(* IEC 61131-3 sources: daoli-st-library/DL_Process (part 15) *)

(* ---- FC_DL_PaddingPickupCalc.st ---- *)
(*
  DL Factory R83 | FC_DL_PaddingPickupCalc
  功能：由轧车前干重与轧后湿重算轧余率，并按克重门幅速度换算带液量。
  开源溯源：无（clean-room 自研，依据公开工艺公式，来源=行业通用公式，许可证=MIT，借鉴点=公式结构）
  规则：R1-R21 全遵守
*)
FUNCTION FC_DL_PaddingPickupCalc : REAL
VAR_INPUT
    fWetMassG : REAL; // 轧后湿重试样质量 [g] / Wet mass after padding [g]
    fDryMassG : REAL; // 轧前干重试样质量 [g] / Dry mass before padding [g]
    fSpeedMpm : REAL; // 轧车线速度 [m/min] / Padder line speed [m/min]
    fWidthM   : REAL; // 织物门幅 [m] / Fabric width [m]
    fGsm      : REAL; // 织物干克重 [g/m²] / Dry grammage [g/m^2]
END_VAR
VAR_OUTPUT
    fPickupPct : REAL; // 轧余率（带液量占干布重）[%] / Wet pickup [%]
    fCarryLpm  : REAL; // 每分钟带液量（密度按 1 kg/L 近似）[L/min] / Liquor carry-over [L/min]
    fCarryKgH  : REAL; // 每小时带液量 [kg/h] / Liquor carry-over [kg/h]
    xValid     : BOOL; // 计算有效性标志 / Calculation validity flag
END_VAR
VAR
    fDryKgMin : REAL; // 每分钟干布质量 [kg/min] / Dry fabric mass per minute [kg/min]
END_VAR
// 出口预置：四出口统一预置（R256）
fPickupPct := 0.0; fCarryLpm := 0.0; fCarryKgH := 0.0; xValid := FALSE;
// 非有限拦截 + 量纲自检 + 湿干重次序闸（R20/R21）
IF NOT (fWetMassG > -1.0E30 AND fWetMassG < 1.0E30) OR NOT (fDryMassG > -1.0E30 AND fDryMassG < 1.0E30) OR NOT (fSpeedMpm > -1.0E30 AND fSpeedMpm < 1.0E30) OR NOT (fWidthM > -1.0E30 AND fWidthM < 1.0E30) OR NOT (fGsm > -1.0E30 AND fGsm < 1.0E30) OR fDryMassG <= 0.0 OR fSpeedMpm <= 0.0 OR fWidthM <= 0.0 OR fGsm <= 0.0 OR fWetMassG < fDryMassG THEN
    FC_DL_PaddingPickupCalc := -1.0; RETURN;   // 哨兵 -1：非有限或量纲/次序越界 / Sentinel -1
END_IF
// 轧余率：(湿重 - 干重) ÷ 干重 × 100，干重分母已零闸（R4/R21）
IF ABS(fDryMassG) > 1.0E-9 THEN                // 干重分母显式零闸 / Explicit zero gate on dry mass
    fPickupPct := (fWetMassG - fDryMassG) / fDryMassG * 100.0; // 轧余率 [%] / Wet pickup [%]
ELSE
    fPickupPct := 0.0;              // 除零防御缺省 [%] / Divide-by-zero default
END_IF
// 每分钟干布质量：g/m² × m × m/min ÷ 1000 = kg/min（m² 与 m 相乘后 g→kg 需除 1000）
fDryKgMin := fGsm * fWidthM * fSpeedMpm / 1000.0;  // 干布质量流率 [kg/min] / Dry mass flow
// 带液量：干布流率 × 轧余率 ÷ 100，密度按 1 kg/L 近似故 kg/min 与 L/min 数值等同
fCarryLpm := fDryKgMin * (fPickupPct / 100.0);     // 每分钟带液 [L/min] / Carry-over [L/min]
fCarryKgH := fCarryLpm * 60.0;                    // 每小时带液 [kg/h] / Carry-over [kg/h]
xValid    := TRUE;                                 // 链路有效 / Chain valid
FC_DL_PaddingPickupCalc := fPickupPct;             // 返回轧余率 [%] / Return wet pickup [%]
END_FUNCTION

(* ---- FC_DL_PaperBasisWeightCalc.st ---- *)
(*
  DL Factory R84 | FC_DL_PaperBasisWeightCalc
  功能：由卷重/幅宽/长度算纸张定量并做水分修正与偏差判定
  开源溯源：无（clean-room 自研，依据公开工艺公式，来源=行业通用公式，许可证=MIT，借鉴点=公式结构）
  规则：R1-R16 全遵守
*)
FUNCTION FC_DL_PaperBasisWeightCalc : REAL
VAR_INPUT
    fRollKg : REAL := 1200.0; // 卷筒重量（含水分） [kg] / roll mass including moisture [kg]
    fWidthM : REAL := 3.5; // 幅宽 [m] / web width [m]
    fLengthM : REAL := 8000.0; // 卷长 [m] / roll length [m]
    fMoistPct : REAL := 7.0; // 成纸水分 [%] / paper moisture [%]
    fTargetGm2 : REAL := 80.0; // 目标定量 [g/m²] / target basis weight [g/m^2]
    fTolPct : REAL := 3.0; // 定量偏差允差 [%] / basis weight tolerance [%]
END_VAR
VAR_OUTPUT
    fDevPct : REAL; // 定量相对偏差 [%] / relative basis weight deviation [%]
    fBoneDryG : REAL; // 绝干质量 [g] / bone dry mass [g]
    xPass : BOOL; // 定量判合格 [-] / basis weight passed [-]
END_VAR
VAR
    fAreaM2 : REAL; // 纸幅面积 [m²] / web area [m^2]
    fBasisGm2 : REAL; // 绝干定量 [g/m²] / bone dry basis weight [g/m^2]
    xValid : BOOL; // 计算有效标志（内部） [-] / internal validity flag [-]
END_VAR

// 段 1｜出口预置（R256）
FC_DL_PaperBasisWeightCalc := -1.0; // 哨兵返回 -1（无效） [-] / sentinel return -1, invalid [-]
fDevPct := 0.0; // 偏差预置零 [%] / deviation preset zero [%]
fBoneDryG := 0.0; // 绝干质量预置零 [g] / bone dry mass preset zero [g]
xPass := FALSE; // 合格位预置 FALSE [-] / pass preset false [-]
xValid := FALSE; // 计算完成前不认结果 [-] / unusable before calculation [-]

// 段 2｜非有限拦截 + 域闸（R4/R20）
IF NOT (fRollKg > -1.0E30 AND fRollKg < 1.0E30) OR NOT (fWidthM > -1.0E30 AND fWidthM < 1.0E30) OR NOT (fLengthM > -1.0E30 AND fLengthM < 1.0E30) THEN
    RETURN; // 卷重/幅宽/卷长任一非有限即拒算 [-] / any non finite roll geometry rejected [-]
END_IF
IF NOT (fMoistPct > -1.0E30 AND fMoistPct < 1.0E30) OR NOT (fTargetGm2 > -1.0E30 AND fTargetGm2 < 1.0E30) OR NOT (fTolPct > -1.0E30 AND fTolPct < 1.0E30) THEN
    RETURN; // 水分/目标定量/允差任一非有限即拒算 [-] / any non finite moisture or target rejected [-]
END_IF
IF fRollKg <= 0.0 OR fWidthM < 1.0E-9 OR fLengthM < 1.0E-9 OR fTargetGm2 < 1.0E-9 OR fTolPct < 0.0 THEN
    RETURN; // 面积与目标定量正域分母闸（防除零） [m, g/m²] / positive denominator gate [m, g/m^2]
END_IF
IF fMoistPct < 0.0 OR fMoistPct >= 100.0 THEN
    RETURN; // 水分开区间域闸 [0,100) [%] / moisture open interval gate [%]
END_IF

// 段 3｜绝干质量与面积
fBoneDryG := (fRollKg * 1000.0) * (1.0 - (fMoistPct / 100.0)); // kg × 1000 g/kg × 无量纲 = g / [kg] × [g/kg] × [-] = [g]
fAreaM2 := fWidthM * fLengthM; // m × m = m² / [m] × [m] = [m^2]
IF fAreaM2 < 1.0E-9 THEN
    RETURN; // 分母闸：面积趋零 [m²] / denominator gate on the area [m^2]
END_IF

// 段 4｜定量与偏差
fBasisGm2 := fBoneDryG / fAreaM2; // g ÷ m² = g/m² / [g] / [m^2] = [g/m^2]
fDevPct := ((fBasisGm2 - fTargetGm2) / fTargetGm2) * 100.0; // (g/m² ÷ g/m²) × 100 = % / [g/m^2] / [g/m^2] × 100 = [%]
IF NOT (fBasisGm2 > -1.0E30 AND fBasisGm2 < 1.0E30) OR NOT (fDevPct > -1.0E30 AND fDevPct < 1.0E30) THEN
    RETURN; // 结果非有限再拦一次 [-] / second finiteness gate on the results [-]
END_IF
xPass := ABS(fDevPct) <= fTolPct; // 偏差绝对值与允差直比 [-] / absolute deviation against the tolerance [-]
xValid := TRUE; // 链路有效 [-] / chain valid [-]
FC_DL_PaperBasisWeightCalc := fBasisGm2; // 返回绝干定量 [g/m²] / return the basis weight [g/m^2]
END_FUNCTION

(* ---- FC_DL_PaperFormationIndexCalc.st ---- *)
(*
  DL Factory R84 | FC_DL_PaperFormationIndexCalc
  功能：由絮聚波长与小尺度方差比估算成形指数（0~1）并按 0.6 判良好
  开源溯源：无（clean-room 自研，依据公开工艺公式，来源=行业通用公式，许可证=MIT，借鉴点=公式结构）
  规则：R1-R16 全遵守
*)
FUNCTION FC_DL_PaperFormationIndexCalc : REAL
VAR_INPUT
    fVarTotal : REAL := 1.0; // 全尺度方差（归一化） [-] / total normalised variance [-]
    fVarSmall : REAL := 0.25; // 小尺度方差分量 [-] / small scale variance component [-]
    fScaleRefMm : REAL := 1.0; // 参考絮聚尺度（像素→mm 标定） [mm] / reference floc scale [mm]
    fLambda0Mm : REAL := 2.0; // 良好成形的特征波长基准 [mm] / reference wavelength of good formation [mm]
    fIdxMin : REAL := 0.6; // 成形指数良好下限 [-] / good formation threshold [-]
END_VAR
VAR_OUTPUT
    fFlocLambda : REAL; // 估算絮聚波长 [mm] / estimated floc wavelength [mm]
    xPass : BOOL; // 成形指数判良好 [-] / formation passed [-]
    xValid : BOOL; // 计算结果有效标志 [-] / calculation valid flag [-]
END_VAR
VAR
    fRatio : REAL; // 全尺度/小尺度方差比 [-] / total to small variance ratio [-]
    fIdxRaw : REAL; // 未钳位成形指数 [-] / unclamped formation index [-]
    fIdx : REAL; // 钳位后成形指数 [-] / clamped formation index [-]
END_VAR

// 段 1｜出口预置（R256）
FC_DL_PaperFormationIndexCalc := -1.0; // 哨兵返回 -1（无效） [-] / sentinel return -1, invalid [-]
fFlocLambda := 0.0; // 絮聚波长预置零 [mm] / floc wavelength preset zero [mm]
xPass := FALSE; // 良好位预置 FALSE [-] / pass preset false [-]
xValid := FALSE; // 计算完成前不认结果 [-] / unusable before calculation [-]

// 段 2｜非有限拦截 + 域闸（R4/R20）
IF NOT (fVarTotal > -1.0E30 AND fVarTotal < 1.0E30) OR NOT (fVarSmall > -1.0E30 AND fVarSmall < 1.0E30) OR NOT (fScaleRefMm > -1.0E30 AND fScaleRefMm < 1.0E30) THEN
    RETURN; // 方差与标定尺度任一非有限即拒算 [-] / any non finite variance or scale rejected [-]
END_IF
IF NOT (fLambda0Mm > -1.0E30 AND fLambda0Mm < 1.0E30) OR NOT (fIdxMin > -1.0E30 AND fIdxMin < 1.0E30) THEN
    RETURN; // 基准波长与门限任一非有限即拒算 [-] / any non finite reference or threshold rejected [-]
END_IF
IF fVarTotal < 0.0 OR fVarSmall < 1.0E-9 OR fScaleRefMm < 1.0E-9 OR fLambda0Mm < 1.0E-9 THEN
    RETURN; // 方差非负 + 小尺度方差/尺度/基准正域分母闸（防除零） [-] / non negative variance and positive denominator gate [-]
END_IF

// 段 3｜方差比与絮聚波长估算（mm × 无量纲 = mm）
fRatio := fVarTotal / fVarSmall; // 无量纲 / [-] = [-] / [-] / [-] = [-]
fFlocLambda := fScaleRefMm * fRatio; // mm × 无量纲 = mm / [mm] × [-] = [mm]
IF NOT (fFlocLambda > -1.0E30 AND fFlocLambda < 1.0E30) THEN
    RETURN; // 结果非有限再拦一次 [-] / second finiteness gate [-]
END_IF

// 段 4｜成形指数 = λ0 / (λ0 + λfloc)，钳位到 0~1
fIdxRaw := fLambda0Mm / (fLambda0Mm + fFlocLambda); // mm ÷ mm = 无量纲 / [mm] / [mm] = [-]
fIdx := fIdxRaw; // 先接未钳位值 [-] / take the raw index [-]
IF fIdx > 1.0 THEN
    fIdx := 1.0; // 上限钳位 [-] / clamp high [-]
END_IF
IF fIdx < 0.0 THEN
    fIdx := 0.0; // 下限钳位（指数物理区间 0~1） [-] / clamp low to the physical range [-]
END_IF

// 段 5｜良好判定与出口
xPass := fIdx >= fIdxMin; // 直比门限，禁浮点等值 [-] / direct compare against the threshold [-]
xValid := TRUE; // 链路有效 [-] / chain valid [-]
FC_DL_PaperFormationIndexCalc := fIdx; // 返回成形指数 [-] / return the formation index [-]
END_FUNCTION

(* ---- FC_DL_PlatingThicknessChargeCalc.st ---- *)
(*
  DL Factory R83 | FC_DL_PlatingThicknessChargeCalc
  功能：按法拉第定律由电流密度、时间与电流效率算镀层厚度并折算电量。
  开源溯源：无（clean-room 自研，依据公开工艺公式，来源=行业通用公式，许可证=MIT，借鉴点=公式结构）
  规则：R1-R21 全遵守
*)
FUNCTION FC_DL_PlatingThicknessChargeCalc : REAL
VAR_INPUT
    fCurrentDens  : REAL; // 阴极电流密度 [A/dm²] / Cathodic current density [A/dm^2]
    fTimeS        : REAL; // 通电时间 [s] / Plating time [s]
    fEffPct       : REAL; // 电流效率（0~100）[%] / Current efficiency [%]
    fEquivMgC     : REAL; // 电化当量 [mg/C] / Electrochemical equivalent [mg/C]
    fMetalDensity : REAL; // 镀层金属密度 [g/cm³] / Deposit density [g/cm^3]
END_VAR
VAR_OUTPUT
    fMassG    : REAL; // 单位面积沉积质量 [g/dm²] / Deposited mass per area [g/dm^2]
    fThickUm  : REAL; // 镀层厚度 [µm] / Deposit thickness [um]
    fChargeAh : REAL; // 单位面积电量 [Ah/dm²] / Charge per area [Ah/dm^2]
    xValid    : BOOL; // 计算有效性标志 / Calculation validity flag
END_VAR
VAR
    fEffK : REAL; // 电流效率归一化系数 [-]/ Normalised efficiency factor
END_VAR
// 出口预置：四出口统一预置（R256）
fMassG := 0.0; fThickUm := 0.0; fChargeAh := 0.0; xValid := FALSE;
// 非有限拦截 + 量纲自检（R20/R21）
IF NOT (fCurrentDens > -1.0E30 AND fCurrentDens < 1.0E30) OR NOT (fTimeS > -1.0E30 AND fTimeS < 1.0E30) OR NOT (fEffPct > -1.0E30 AND fEffPct < 1.0E30) OR NOT (fEquivMgC > -1.0E30 AND fEquivMgC < 1.0E30) OR NOT (fMetalDensity > -1.0E30 AND fMetalDensity < 1.0E30) OR fCurrentDens < 0.0 OR fTimeS < 0.0 OR fEquivMgC <= 0.0 OR fMetalDensity <= 0.0 THEN
    FC_DL_PlatingThicknessChargeCalc := -1.0; RETURN; // 哨兵 -1：非有限或量纲越界 / Sentinel -1
END_IF
// 电流效率域闸：0~100% 之外钳位（效率不可能超 100）
IF fEffPct < 0.0 THEN
    fEffK := 0.0;                   // 效率零下限 [-] / Efficiency lower bound zero
ELSIF fEffPct > 100.0 THEN
    fEffK := 1.0;                   // 效率满上限 [-] / Efficiency upper bound unity
ELSE
    fEffK := fEffPct / 100.0;       // 归一化效率 [-] / Normalised efficiency
END_IF
// 沉积质量：mg/C ÷ 1000 = g/C；g/C × A/dm² × s = g/dm²（量纲自洽：C = A·s）
fMassG := (fEquivMgC / 1000.0) * fEffK * fCurrentDens * fTimeS; // 单位面积质量 [g/dm²]
// 厚度：1 dm² = 100 cm²，故 µm = 100 × (g/dm²) ÷ (g/cm³)，密度分母显式零闸（R4/R21）
IF ABS(fMetalDensity) > 1.0E-9 THEN            // 密度分母显式零闸 / Explicit zero gate on density
    fThickUm := 100.0 * fMassG / fMetalDensity; // 镀层厚度 [µm] / Deposit thickness [um]
ELSE
    fThickUm := 0.0;                // 除零防御缺省 [µm] / Divide-by-zero default
END_IF
// 电量：A/dm² × s ÷ 3600 = Ah/dm²（s→h 换算常数 3600）
fChargeAh := fCurrentDens * fTimeS / 3600.0;   // 单位面积电量 [Ah/dm²] / Charge per area
xValid    := TRUE;                             // 链路有效 / Chain valid
FC_DL_PlatingThicknessChargeCalc := fThickUm;  // 返回镀层厚度 [µm] / Return deposit thickness
END_FUNCTION

(* ---- FC_DL_PolymerDoseCalc.st ---- *)
(*
  道莅工业代码库 / Daoli Industrial ST Library
  组件: FC_DL_PolymerDoseCalc
  分类: DL_Process
  开源溯源: 无（clean-room 工程公式自研；参考公开工艺计算公式，未复制任何受版权保护代码）
  许可证: 本项目自有 (MIT)
  功能: PAM 絮凝剂按干固体单耗折算质量投加量与母液体积投加量
  近似说明: 母液按「1 kg 溶液 ≈ 1 L」折算（浓度 ≤1% 时误差 <1%），已在公式处声明
*)
FUNCTION FC_DL_PolymerDoseCalc : BOOL
VAR_INPUT
    rDsKgH : REAL; // 干固体处理量 [kg/h] / dry solids throughput
    rDoseKgT : REAL; // PAM 单耗（每吨干固体）[kg/t] / polymer dose per tonne of dry solids
    rStockPct : REAL; // 母液配制浓度 [%] / stock solution concentration
END_VAR
VAR_OUTPUT
    rPolyKgH : REAL; // PAM 纯质投加量 [kg/h] / neat polymer mass flow
    rPolyLh : REAL; // PAM 母液体积投加量 [L/h] / stock solution volumetric flow
    bValid : BOOL; // 结果有效位 [-] / result valid flag
    iErrCode : INT; // 事件码 0=正常 1=母液浓度超域 2=单耗为负 3=结果非有限 / event code
END_VAR
VAR CONSTANT
    rKgPerT : REAL := 1000.0; // 每吨公斤数 [kg/t] / kilograms per tonne
    rPctToFrac : REAL := 0.01; // 百分数转小数系数 [-]/[%] / percent to fraction factor
END_VAR
VAR
    rDsTh : REAL; // 干固体处理量 [t/h] / dry solids in tonnes per hour
    rPolyRaw : REAL; // 未限幅纯质投加 [kg/h] / unchecked neat polymer flow
    rStockFrac : REAL; // 母液质量分数 [-] / stock mass fraction
END_VAR

    // —— 段 0：全路径预清 —— //
    rDsTh := 0.0;
    rPolyRaw := 0.0;
    rStockFrac := 0.0;
    rPolyKgH := 0.0;
    rPolyLh := 0.0;
    bValid := FALSE;
    iErrCode := 0;
    FC_DL_PolymerDoseCalc := FALSE;
    // —— 段 1：母液浓度域闸 (0, 100]% 兼分母闸 —— //
    IF (rStockPct <= 0.0) OR (rStockPct > 100.0) THEN
        iErrCode := 1; // 母液浓度超域，体积流量无定义 / stock concentration out of domain
        RETURN;
    END_IF;
    IF rDoseKgT < 0.0 THEN
        iErrCode := 2; // 单耗为负，拒绝换算 / negative dose rejected
        RETURN;
    END_IF;
    // —— 段 2：量纲链 (kg/h)/(kg/t) = t/h；(t/h)*(kg/t) = kg/h —— //
    rDsTh := rDsKgH / rKgPerT; // 干固体 [t/h] / dry solids in t/h
    rPolyRaw := rDsTh * rDoseKgT; // 纯质 PAM [kg/h] / neat polymer flow
    IF ABS(rPolyRaw) > 1.0E15 THEN
        iErrCode := 3; // 结果非有限，强制归零 / non-finite result, forced to zero
        RETURN;
    END_IF;
    IF rPolyRaw < 0.0 THEN
        rPolyKgH := 0.0; // 负干固体防御 / negative dry solids guard
    ELSE
        rPolyKgH := rPolyRaw;
    END_IF;
    // —— 段 3：母液体积 = 纯质量 / 质量分数（1 kg 溶液 ≈ 1 L 近似） —— //
    rStockFrac := rStockPct * rPctToFrac; // 质量分数 [-] / stock mass fraction
    rPolyLh := rPolyKgH / rStockFrac; // 母液体积 [L/h] / stock volumetric flow
    IF ABS(rPolyLh) > 1.0E15 THEN
        rPolyLh := 0.0;
        iErrCode := 3; // 结果非有限，强制归零 / non-finite result, forced to zero
        RETURN;
    END_IF;
    bValid := TRUE;
    FC_DL_PolymerDoseCalc := TRUE;
END_FUNCTION

(* ---- FC_DL_PotlineAluminaFeedRateCalc.st ---- *)
// FC_DL_PotlineAluminaFeedRateCalc v1.0.0
// 开源溯源：clean-room 自研（族 DL_Process，ST 生态实测 0 命中，无外部代码引入）
(*
  功能: 产铝率 = I[kA]·0.3355·CE/100 [kg/h]（0.3355 为铝电化学当量），
        Al2O3 理论量 = 产铝·1.889，下料率 = 理论量/(1 − 损耗率/100)。
  邻件/码位: 与 FC_DL_PotlineCurrentEfficiencyCalc 互为逆过程（本件由 CE 正算产物与下料）；
             16#0002_9212 = 非有限、CE 越界或损耗率 ≥ 100% 拒收。
*)
FUNCTION FC_DL_PotlineAluminaFeedRateCalc : REAL
VAR_INPUT
    fCurrentKA  : REAL := 400.0;    // 系列电流 [kA]，域 > 0 / Line current [kA]
    fCE         : REAL := 93.0;     // 电流效率 [%]，域 (0, 100] / Current efficiency [%]
    fLossRatio  : REAL := 2.0;      // 氧化铝损耗率 [%]，域 [0, 100) / Alumina loss ratio [%]
END_VAR
VAR_OUTPUT
    fAlRate      : REAL;            // 产铝速率 [kg/h] / Aluminium production rate [kg/h]
    fAluminaRate : REAL;            // 氧化铝下料率 [kg/h] / Alumina feed rate [kg/h]
    bValid       : BOOL;            // 结果有效回执 [-] / Result validity receipt
    uErrorId     : UDINT;           // 事件码，0 = 无事件 / Event code
END_VAR
VAR
    fLossFrac : REAL := 0.0;        // 损耗率小数 [-] / Loss ratio as fraction [-]
END_VAR
// 段 0：全路径出口安全缺省 / Safe defaults on all outlets
fAlRate := 0.0;                 // 产铝速率缺省零 / Production rate default zero
fAluminaRate := 0.0;            // 下料率缺省零 / Feed rate default zero
bValid := FALSE;                // 有效回执预清 / Validity preset clear
uErrorId := 16#0000;            // 事件码预清 / Event code preset clear
FC_DL_PotlineAluminaFeedRateCalc := 0.0;    // 返回值缺省零（镜像产铝）/ Return default zero
// 段 1：非有限闸（三入参全枚举）/ Non-finite gate over all inputs
IF (fCurrentKA <> fCurrentKA) OR (fCE <> fCE) OR (fLossRatio <> fLossRatio)
   OR (ABS(fCurrentKA) >= 3.0E38) OR (ABS(fCE) >= 3.0E38) OR (ABS(fLossRatio) >= 3.0E38) THEN
    uErrorId := 16#0002_9212;   // 入参非有限拒收 / Non-finite input reject
    RETURN;
END_IF
// 段 2：域闸（电流正 / CE 区间 / 损耗率上界防除零，R4）/ Domain gate
IF fCurrentKA <= 1.0E-6 THEN
    uErrorId := 16#0002_9212;   // 电流非正 / Non-positive current
    RETURN;
END_IF
IF (fCE <= 0.0) OR (fCE > 100.0) THEN
    uErrorId := 16#0002_9212;   // 电流效率越界 / Current efficiency out of range
    RETURN;
END_IF
IF (fLossRatio < 0.0) OR (fLossRatio >= 100.0) THEN
    uErrorId := 16#0002_9212;   // 损耗率越界（分母 1−loss 近零）/ Loss ratio out of range
    RETURN;
END_IF
// 段 3：主计算（产物 → 理论氧化铝 → 损耗补正下料）/ Main computation
fAlRate := fCurrentKA * 0.3355 * fCE / 100.0;                   // 产铝 = I·当量·CE / Production rate
fLossFrac := fLossRatio / 100.0;                                // 损耗率转小数 / Loss as fraction
fAluminaRate := fAlRate * 1.889 / (1.0 - fLossFrac);            // 损耗补正下料 / Loss-compensated feed
// 段 4：出口闸（双输出非有限复核 + 非负复核）/ Outlet gate
IF (fAlRate <> fAlRate) OR (fAluminaRate <> fAluminaRate)
   OR (ABS(fAlRate) >= 3.0E38) OR (ABS(fAluminaRate) >= 3.0E38)
   OR (fAlRate < 0.0) OR (fAluminaRate < 0.0) THEN
    fAlRate := 0.0;             // 复核失败回缺省 / Fallback on recheck failure
    fAluminaRate := 0.0;        // 复核失败回缺省 / Fallback on recheck failure
    uErrorId := 16#0002_9212;   // 出口复核拒收 / Output recheck reject
    RETURN;
END_IF
bValid := TRUE;                 // 有效回执 / Validity receipt
FC_DL_PotlineAluminaFeedRateCalc := fAlRate;    // 返回值镜像产铝速率 / Return mirrors rate
END_FUNCTION

(* ---- FC_DL_PotlineAnodeEffectEnergyCalc.st ---- *)
// FC_DL_PotlineAnodeEffectEnergyCalc v1.0.0
// 开源溯源：clean-room 自研（族 DL_Process，ST 生态实测 0 命中，无外部代码引入）
(*
  功能: 效应能耗核算：单次能耗 = V·I[kA]·t[min]/60 [kWh]（kA·V·min/60 = kWh），
        日能耗 = 单次 × 日次数；效应系数按「次/槽日」出口（统计窗为 24 h 槽日）。
  邻件/码位: 与 FC_DL_PotlineCellVoltageBudgetCalc 分域（效应附加电耗 vs 正常槽电压）；
             16#0002_9213 = 非有限、电压/电流/时长非正或次数为负拒收。
*)
FUNCTION FC_DL_PotlineAnodeEffectEnergyCalc : REAL
VAR_INPUT
    fEffectVoltage : REAL := 8.0;   // 效应净增电压 [V]，域 > 0 / Net effect voltage [V]
    fLineCurrentKA : REAL := 400.0; // 系列电流 [kA]，域 > 0 / Line current [kA]
    fEffectMin     : REAL := 3.0;   // 单次效应时长 [min]，域 > 0 / Effect duration [min]
    fEffectsPerDay : REAL := 0.5;   // 日效应次数 [次/日]，域 >= 0 / Effects per day [count/day]
END_VAR
VAR_OUTPUT
    fEnergyPerEffect   : REAL;      // 单次效应能耗 [kWh] / Energy per effect [kWh]
    fEffectCoefficient : REAL;      // 效应系数 [次/槽日] / Effect coefficient [count/pot-day]
    fDailyEnergy       : REAL;      // 日效应能耗 [kWh/日] / Daily energy [kWh/day]
    bValid             : BOOL;      // 结果有效回执 [-] / Result validity receipt
    uErrorId           : UDINT;     // 事件码，0 = 无事件 / Event code
END_VAR
// 段 0：全路径出口安全缺省 / Safe defaults on all outlets
fEnergyPerEffect := 0.0;            // 单次能耗缺省零 / Per-effect default zero
fEffectCoefficient := 0.0;          // 效应系数缺省零 / Coefficient default zero
fDailyEnergy := 0.0;                // 日能耗缺省零 / Daily energy default zero
bValid := FALSE;                    // 有效回执预清 / Validity preset clear
uErrorId := 16#0000;                // 事件码预清 / Event code preset clear
FC_DL_PotlineAnodeEffectEnergyCalc := 0.0;  // 返回值缺省零（镜像单次能耗）/ Return default zero
// 段 1：非有限闸（四入参全枚举）/ Non-finite gate over all inputs
IF (fEffectVoltage <> fEffectVoltage) OR (fLineCurrentKA <> fLineCurrentKA)
   OR (fEffectMin <> fEffectMin) OR (fEffectsPerDay <> fEffectsPerDay)
   OR (ABS(fEffectVoltage) >= 3.0E38) OR (ABS(fLineCurrentKA) >= 3.0E38)
   OR (ABS(fEffectMin) >= 3.0E38) OR (ABS(fEffectsPerDay) >= 3.0E38) THEN
    uErrorId := 16#0002_9213;   // 入参非有限拒收 / Non-finite input reject
    RETURN;
END_IF
// 段 2：域闸（电压/电流/时长为正 + 次数非负）/ Domain gate
IF (fEffectVoltage <= 0.0) OR (fLineCurrentKA <= 1.0E-6) OR (fEffectMin <= 1.0E-6) THEN
    uErrorId := 16#0002_9213;   // 电压、电流或时长非正 / Non-positive voltage, current or duration
    RETURN;
END_IF
IF fEffectsPerDay < 0.0 THEN
    uErrorId := 16#0002_9213;   // 效应次数为负 / Negative effect count
    RETURN;
END_IF
// 段 3：主计算（单次能耗 → 效应系数 → 日能耗）/ Main computation
fEnergyPerEffect := fEffectVoltage * fLineCurrentKA * fEffectMin / 60.0;    // V·I·t/60 [kWh] / Per effect
fEffectCoefficient := fEffectsPerDay;                           // 24 h 槽日内即次数本身 / Count over 24h
fDailyEnergy := fEnergyPerEffect * fEffectsPerDay;              // 日能耗 / Daily energy
// 段 4：出口闸（三输出非有限复核 + 非负复核）/ Outlet gate
IF (fEnergyPerEffect <> fEnergyPerEffect) OR (fEffectCoefficient <> fEffectCoefficient)
   OR (fDailyEnergy <> fDailyEnergy)
   OR (ABS(fEnergyPerEffect) >= 3.0E38) OR (ABS(fEffectCoefficient) >= 3.0E38)
   OR (ABS(fDailyEnergy) >= 3.0E38) THEN
    fEnergyPerEffect := 0.0;        // 复核失败回缺省 / Fallback on recheck failure
    fEffectCoefficient := 0.0;      // 复核失败回缺省 / Fallback on recheck failure
    fDailyEnergy := 0.0;            // 复核失败回缺省 / Fallback on recheck failure
    uErrorId := 16#0002_9213;       // 出口非有限拒收 / Output non-finite reject
    RETURN;
END_IF
bValid := TRUE;                     // 有效回执 / Validity receipt
FC_DL_PotlineAnodeEffectEnergyCalc := fEnergyPerEffect;     // 返回值镜像单次能耗 / Return mirrors
END_FUNCTION

(* ---- FC_DL_PotlineBathRatioCalc.st ---- *)
// FC_DL_PotlineBathRatioCalc v1.0.0
// 开源溯源：clean-room 自研（族 DL_Process，ST 生态实测 0 命中，无外部代码引入）
(*
  功能: 电解质分子比 CR = (wNaF/41.99)/(wAlF3/83.97)（41.99/83.97 为 NaF/AlF3 摩尔质量），
        过剩 AlF3 = wAlF3 − (wNaF·83.97/41.99)/2 [%]。
  邻件/码位: 与 FC_DL_PotlineBathTempDeviationCalc 构成化验→热状态链（本件出 CR）；
             16#0002_9211 = 非有限、AlF3 过低、成分和超 100% 或 CR 出 1.5~3.5 拒收。
*)
FUNCTION FC_DL_PotlineBathRatioCalc : REAL
VAR_INPUT
    fNaFWt  : REAL := 45.0;     // NaF 质量分数 [%] / NaF mass fraction [%]
    fAlF3Wt : REAL := 40.0;     // AlF3 质量分数 [%]，域 > 0.5 / AlF3 mass fraction [%]
    fCaF2Wt : REAL := 5.0;      // CaF2 质量分数 [%] / CaF2 mass fraction [%]
END_VAR
VAR_OUTPUT
    fCryoliteRatio : REAL;      // 分子比 CR [-]，典型 2.2~2.6 / Cryolite ratio [-]
    fExcessAlF3    : REAL;      // 过剩 AlF3 [%] / Excess AlF3 [%]
    bValid         : BOOL;      // 结果有效回执 [-] / Result validity receipt
    uErrorId       : UDINT;     // 事件码，0 = 无事件 / Event code
END_VAR
VAR
    fMolNaF  : REAL := 0.0;     // NaF 摩尔相对量 [mol] / NaF mole amount [mol]
    fMolAlF3 : REAL := 0.0;     // AlF3 摩尔相对量 [mol] / AlF3 mole amount [mol]
END_VAR
// 段 0：全路径出口安全缺省 / Safe defaults on all outlets
fCryoliteRatio := 0.0;          // 分子比缺省零 / Ratio default zero
fExcessAlF3 := 0.0;             // 过剩 AlF3 缺省零 / Excess default zero
bValid := FALSE;                // 有效回执预清 / Validity preset clear
uErrorId := 16#0000;            // 事件码预清 / Event code preset clear
FC_DL_PotlineBathRatioCalc := 0.0;      // 返回值缺省零（镜像 CR）/ Return default zero
// 段 1：非有限闸（三入参全枚举）/ Non-finite gate over all inputs
IF (fNaFWt <> fNaFWt) OR (fAlF3Wt <> fAlF3Wt) OR (fCaF2Wt <> fCaF2Wt)
   OR (ABS(fNaFWt) >= 3.0E38) OR (ABS(fAlF3Wt) >= 3.0E38) OR (ABS(fCaF2Wt) >= 3.0E38) THEN
    uErrorId := 16#0002_9211;   // 入参非有限拒收 / Non-finite input reject
    RETURN;
END_IF
// 段 2：域闸（AlF3 下界防除零 + 组分非负 + 成分和上界，R4）/ Domain gate
IF (fNaFWt < 0.0) OR (fCaF2Wt < 0.0) OR (fAlF3Wt <= 0.5) THEN
    uErrorId := 16#0002_9211;   // 负组分或 AlF3 过低（分母近零）/ Negative or too-low AlF3
    RETURN;
END_IF
IF (fNaFWt + fAlF3Wt + fCaF2Wt) > 100.0 THEN
    uErrorId := 16#0002_9211;   // 成分和超 100%，化验数据非法 / Sum exceeds 100 percent
    RETURN;
END_IF
// 段 3：主计算（摩尔比 + 过剩 AlF3）/ Main computation
fMolNaF := fNaFWt / 41.99;                                      // NaF 摩尔相对量 / NaF mole amount
fMolAlF3 := fAlF3Wt / 83.97;                                    // AlF3 摩尔相对量 / AlF3 mole amount
fCryoliteRatio := fMolNaF / fMolAlF3;                           // CR = nNaF/nAlF3 / Cryolite ratio
// 过剩 AlF3 基准为冰晶石 CR=3（Na3AlF6 即 3NaF·AlF3），故除以 3 而非 2
// 说明（R92-修正）：早期版本除 2，致纯冰晶石组份（CR=3）输出 −20%，符号与量级双错
fExcessAlF3 := fAlF3Wt - (fNaFWt * 83.97 / 41.99) / 3.0;        // 过剩 AlF3 [%] / Excess AlF3
// 段 4：出口闸（非有限复核 + CR 工艺窗判定）/ Outlet gate
IF (fCryoliteRatio <> fCryoliteRatio) OR (fExcessAlF3 <> fExcessAlF3)
   OR (ABS(fCryoliteRatio) >= 3.0E38) OR (ABS(fExcessAlF3) >= 3.0E38) THEN
    fCryoliteRatio := 0.0;      // 复核失败回缺省 / Fallback on recheck failure
    fExcessAlF3 := 0.0;         // 复核失败回缺省 / Fallback on recheck failure
    uErrorId := 16#0002_9211;   // 出口非有限拒收 / Output non-finite reject
    RETURN;
END_IF
IF (fCryoliteRatio < 1.5) OR (fCryoliteRatio > 3.5) THEN
    uErrorId := 16#0002_9211;   // 信息级：CR 出工艺窗 / Info: ratio out of window
    RETURN;                     // bValid 保持 FALSE / Validity stays false
END_IF
bValid := TRUE;                 // 有效回执 / Validity receipt
FC_DL_PotlineBathRatioCalc := fCryoliteRatio;   // 返回值镜像 CR / Return mirrors ratio
END_FUNCTION

(* ---- FC_DL_PotlineBathTempDeviationCalc.st ---- *)
// FC_DL_PotlineBathTempDeviationCalc v1.0.0
// 开源溯源：clean-room 自研（族 DL_Process，ST 生态实测 0 命中，无外部代码引入）
(*
  功能: 初晶温度简化线性工程近似式（非相图严格解）：
        T_liq = 961.0 − 12.5·(CR − 2.0) − 3.5·(CaF2/100·100)/8.0 − 2.0·(MgF2/8.0)，
        过热度 = 槽温 − 初晶温度，> 12 °C 置 bOverheat。961.0 为 CR=2.0 无添加剂的基准初晶温度。
  邻件/码位: 与 FC_DL_PotlineBathRatioCalc 串联（前件出 CR）；与 FC_DL_PotlineMetalLevelCalc 同族不同域；
             16#0002_9216 = 非有限、CR 出 1.5~3.5 或添加剂为负拒收。
*)
FUNCTION FC_DL_PotlineBathTempDeviationCalc : REAL
VAR_INPUT
    fBathTemp : REAL := 960.0;      // 槽温（电解质温度）[°C] / Bath temperature [degC]
    fCR       : REAL := 2.30;       // 分子比 CR [-]，域 1.5~3.5 / Cryolite ratio [-]
    fCaF2     : REAL := 5.0;        // CaF2 质量分数 [%] / CaF2 mass fraction [%]
    fMgF2     : REAL := 0.5;        // MgF2 质量分数 [%] / MgF2 mass fraction [%]
END_VAR
VAR_OUTPUT
    fLiquidus  : REAL;              // 初晶温度 [°C] / Liquidus temperature [degC]
    fSuperheat : REAL;              // 过热度 [°C] / Superheat [degC]
    bOverheat  : BOOL;              // 过热告警（> 12 °C）[-] / Overheat alarm flag
    bValid     : BOOL;              // 结果有效回执 [-] / Result validity receipt
    uErrorId   : UDINT;             // 事件码，0 = 无事件 / Event code
END_VAR
// 段 0：全路径出口安全缺省 / Safe defaults on all outlets
fLiquidus := 0.0;               // 初晶温度缺省零 / Liquidus default zero
fSuperheat := 0.0;              // 过热度缺省零 / Superheat default zero
bOverheat := FALSE;             // 过热告警预清 / Overheat preset clear
bValid := FALSE;                // 有效回执预清 / Validity preset clear
uErrorId := 16#0000;            // 事件码预清 / Event code preset clear
FC_DL_PotlineBathTempDeviationCalc := 0.0;  // 返回值缺省零（镜像过热度）/ Return default zero
// 段 1：非有限闸（四入参全枚举）/ Non-finite gate over all inputs
IF (fBathTemp <> fBathTemp) OR (fCR <> fCR) OR (fCaF2 <> fCaF2) OR (fMgF2 <> fMgF2)
   OR (ABS(fBathTemp) >= 3.0E38) OR (ABS(fCR) >= 3.0E38)
   OR (ABS(fCaF2) >= 3.0E38) OR (ABS(fMgF2) >= 3.0E38) THEN
    uErrorId := 16#0002_9216;   // 入参非有限拒收 / Non-finite input reject
    RETURN;
END_IF
// 段 2：域闸（CR 工艺区间，防线性式外推失真 + 添加剂非负）/ Domain gate
IF (fCR < 1.5) OR (fCR > 3.5) THEN
    uErrorId := 16#0002_9216;   // CR 出 1.5~3.5，线性式不适用 / CR out of valid range
    RETURN;
END_IF
IF (fCaF2 < 0.0) OR (fMgF2 < 0.0) THEN
    uErrorId := 16#0002_9216;   // 添加剂质量分数为负 / Negative additive fraction
    RETURN;
END_IF
// 段 3：主计算（线性初晶温度式 + 过热度；CaF2 保留原式形态）/ Main computation
fLiquidus := 961.0
           - 12.5 * (fCR - 2.0)
           - 3.5 * (fCaF2 / 100.0 * 100.0) / 8.0
           - 2.0 * (fMgF2 / 8.0);                               // 初晶温度线性近似 / Linear liquidus
fSuperheat := fBathTemp - fLiquidus;                            // 过热度 = 槽温 − 初晶 / Superheat
IF fSuperheat > 12.0 THEN
    bOverheat := TRUE;          // 过 12 °C 告警 / Alarm above 12 degC
END_IF
// 段 4：出口闸（双输出非有限复核）/ Outlet gate
IF (fLiquidus <> fLiquidus) OR (fSuperheat <> fSuperheat)
   OR (ABS(fLiquidus) >= 3.0E38) OR (ABS(fSuperheat) >= 3.0E38) THEN
    fLiquidus := 0.0;           // 复核失败回缺省 / Fallback on recheck failure
    fSuperheat := 0.0;          // 复核失败回缺省 / Fallback on recheck failure
    bOverheat := FALSE;         // 复核失败清告警 / Clear alarm on recheck failure
    uErrorId := 16#0002_9216;   // 出口非有限拒收 / Output non-finite reject
    RETURN;
END_IF
bValid := TRUE;                 // 有效回执 / Validity receipt
FC_DL_PotlineBathTempDeviationCalc := fSuperheat;   // 返回值镜像过热度 / Return mirrors superheat
END_FUNCTION

(* ---- FC_DL_PotlineBusbarShuntCalc.st ---- *)
// FC_DL_PotlineBusbarShuntCalc v1.0.0
// 开源溯源：clean-room 自研（族 DL_Process，ST 生态实测 0 命中，无外部代码引入）
(*
  功能: 母线并联支路分流：分流比 = R_other/(R_branch + R_other)，支路电流 = 总电流 × 分流比；
        两电阻同为 µΩ 量纲，比值无量纲故不换算。用于母线搭接电阻劣化诊断。
  邻件/码位: 与 FC_DL_PotlineCellVoltageBudgetCalc 层次不同（槽外母线分流 vs 槽内压降）；
             16#0002_9218 = 非有限、总电流非正或任一电阻非正拒收。
*)
FUNCTION FC_DL_PotlineBusbarShuntCalc : REAL
VAR_INPUT
    fTotalCurrent : REAL := 400.0;  // 总电流 [kA]，域 > 0 / Total current [kA]
    fBranchRes    : REAL := 10.0;   // 本支路电阻 [µΩ]，域 > 0 / Branch resistance [uOhm]
    fOtherRes     : REAL := 12.0;   // 其余并联等效电阻 [µΩ]，域 > 0 / Other resistance [uOhm]
END_VAR
VAR_OUTPUT
    fBranchCurrent : REAL;          // 本支路电流 [kA] / Branch current [kA]
    fShuntRatio    : REAL;          // 分流比 [-] / Shunt ratio [-]
    bValid         : BOOL;          // 结果有效回执 [-] / Result validity receipt
    uErrorId       : UDINT;         // 事件码，0 = 无事件 / Event code
END_VAR
VAR
    fResSum : REAL := 0.0;          // 电阻和 [µΩ] / Resistance sum [uOhm]
END_VAR
// 段 0：全路径出口安全缺省 / Safe defaults on all outlets
fBranchCurrent := 0.0;              // 支路电流缺省零 / Branch current default zero
fShuntRatio := 0.0;                 // 分流比缺省零 / Shunt ratio default zero
bValid := FALSE;                    // 有效回执预清 / Validity preset clear
uErrorId := 16#0000;                // 事件码预清 / Event code preset clear
FC_DL_PotlineBusbarShuntCalc := 0.0;        // 返回值缺省零（镜像支路电流）/ Return default zero
// 段 1：非有限闸（三入参全枚举）/ Non-finite gate over all inputs
IF (fTotalCurrent <> fTotalCurrent) OR (fBranchRes <> fBranchRes) OR (fOtherRes <> fOtherRes)
   OR (ABS(fTotalCurrent) >= 3.0E38) OR (ABS(fBranchRes) >= 3.0E38) OR (ABS(fOtherRes) >= 3.0E38) THEN
    uErrorId := 16#0002_9218;   // 入参非有限拒收 / Non-finite input reject
    RETURN;
END_IF
// 段 2：域闸（总电流为正 + 两电阻为正，分母非零，R4）/ Domain gate
IF fTotalCurrent <= 1.0E-6 THEN
    uErrorId := 16#0002_9218;   // 总电流非正 / Non-positive total current
    RETURN;
END_IF
IF (fBranchRes <= 0.0) OR (fOtherRes <= 0.0) THEN
    uErrorId := 16#0002_9218;   // 支路或并联电阻非正 / Non-positive resistance
    RETURN;
END_IF
// 段 3：主计算（分流比 → 支路电流）/ Main computation
fResSum := fBranchRes + fOtherRes;                              // 电阻和 / Resistance sum
fShuntRatio := fOtherRes / fResSum;                             // 分流比 / Shunt ratio
fBranchCurrent := fTotalCurrent * fShuntRatio;                   // 支路电流 / Branch current
// 段 4：出口闸（非有限复核 + 分流比区间复核）/ Outlet gate
IF (fBranchCurrent <> fBranchCurrent) OR (fShuntRatio <> fShuntRatio)
   OR (ABS(fBranchCurrent) >= 3.0E38) OR (ABS(fShuntRatio) >= 3.0E38)
   OR (fShuntRatio <= 0.0) OR (fShuntRatio >= 1.0) THEN
    fBranchCurrent := 0.0;      // 复核失败回缺省 / Fallback on recheck failure
    fShuntRatio := 0.0;         // 复核失败回缺省 / Fallback on recheck failure
    uErrorId := 16#0002_9218;   // 出口复核拒收 / Output recheck reject
    RETURN;
END_IF
bValid := TRUE;                 // 有效回执 / Validity receipt
FC_DL_PotlineBusbarShuntCalc := fBranchCurrent;     // 返回值镜像支路电流 / Return mirrors current
END_FUNCTION

(* ---- FC_DL_PotlineCellVoltageBudgetCalc.st ---- *)
// FC_DL_PotlineCellVoltageBudgetCalc v1.0.0
// 开源溯源：clean-room 自研（族 DL_Process，ST 生态实测 0 命中，无外部代码引入）
(*
  功能: 槽电压预算：Rtot = (R_bath + R_anode)·1e-6 [Ω]，I = I[kA]·1000 [A]，
        欧姆压降 = I·Rtot，槽电压 = 反电动势 + 浓差 + 活化 + 欧姆压降；
        结果出 2.0~8.0 V 工艺窗置 bValid FALSE（工艺异常域，非计算错误）。
  邻件/码位: 与 FC_DL_PotlineAnodeEffectEnergyCalc 分域（正常电压分解 vs 效应附加电耗）；
             16#0002_9214 = 非有限、电阻为负或电流非正或电压出工艺窗。
*)
FUNCTION FC_DL_PotlineCellVoltageBudgetCalc : REAL
VAR_INPUT
    fRevEMF    : REAL := 1.20;      // 反电动势 [V] / Reversible EMF [V]
    fConcOver  : REAL := 0.10;      // 浓差过电位 [V] / Concentration overpotential [V]
    fActOver   : REAL := 0.35;      // 活化过电位 [V] / Activation overpotential [V]
    fBathRes   : REAL := 3.0;       // 电解质电阻 [µΩ]，域 >= 0 / Bath resistance [uOhm]
    fAnodeRes  : REAL := 1.5;       // 阳极气泡电阻 [µΩ]，域 >= 0 / Anode bubble resistance [uOhm]
    fCurrentKA : REAL := 400.0;     // 系列电流 [kA]，域 > 0 / Line current [kA]
END_VAR
VAR_OUTPUT
    fCellVoltage : REAL;            // 槽电压 [V]，工艺域 2.0~8.0 / Cell voltage [V]
    fOhmicDrop   : REAL;            // 欧姆压降 [V] / Ohmic voltage drop [V]
    bValid       : BOOL;            // 结果有效回执 [-] / Result validity receipt
    uErrorId     : UDINT;           // 事件码，0 = 无事件 / Event code
END_VAR
VAR
    fResTotal : REAL := 0.0;        // 总电阻 [Ω] / Total resistance [Ohm]
    fCurrentA : REAL := 0.0;        // 电流 [A] / Current [A]
END_VAR
// 段 0：全路径出口安全缺省 / Safe defaults on all outlets
fCellVoltage := 0.0;                // 槽电压缺省零 / Cell voltage default zero
fOhmicDrop := 0.0;                  // 欧姆压降缺省零 / Ohmic drop default zero
bValid := FALSE;                    // 有效回执预清 / Validity preset clear
uErrorId := 16#0000;                // 事件码预清 / Event code preset clear
FC_DL_PotlineCellVoltageBudgetCalc := 0.0;  // 返回值缺省零（镜像槽电压）/ Return default zero
// 段 1：非有限闸（六入参全枚举）/ Non-finite gate over all inputs
IF (fRevEMF <> fRevEMF) OR (fConcOver <> fConcOver) OR (fActOver <> fActOver)
   OR (fBathRes <> fBathRes) OR (fAnodeRes <> fAnodeRes) OR (fCurrentKA <> fCurrentKA)
   OR (ABS(fRevEMF) >= 3.0E38) OR (ABS(fConcOver) >= 3.0E38) OR (ABS(fActOver) >= 3.0E38)
   OR (ABS(fBathRes) >= 3.0E38) OR (ABS(fAnodeRes) >= 3.0E38) OR (ABS(fCurrentKA) >= 3.0E38) THEN
    uErrorId := 16#0002_9214;   // 入参非有限拒收 / Non-finite input reject
    RETURN;
END_IF
// 段 2：域闸（电阻非负 + 电流为正）/ Domain gate
IF (fBathRes < 0.0) OR (fAnodeRes < 0.0) THEN
    uErrorId := 16#0002_9214;   // 电阻为负，物理非法 / Negative resistance
    RETURN;
END_IF
IF fCurrentKA <= 1.0E-6 THEN
    uErrorId := 16#0002_9214;   // 电流非正 / Non-positive current
    RETURN;
END_IF
// 段 3：主计算（电阻链 → 欧姆压降 → 电压预算）/ Main computation
fResTotal := (fBathRes + fAnodeRes) * 1.0E-6;                   // 总电阻 [Ω] / Total resistance
fCurrentA := fCurrentKA * 1000.0;                               // 电流 [A] / Current in amperes
fOhmicDrop := fCurrentA * fResTotal;                            // 欧姆压降 I·R [V] / Ohmic drop
fCellVoltage := fRevEMF + fConcOver + fActOver + fOhmicDrop;    // 槽电压预算 / Cell voltage budget
// 段 4：出口闸（非有限复核 + 2.0~8.0 V 工艺域判定）/ Outlet gate
IF (fCellVoltage <> fCellVoltage) OR (fOhmicDrop <> fOhmicDrop)
   OR (ABS(fCellVoltage) >= 3.0E38) OR (ABS(fOhmicDrop) >= 3.0E38) THEN
    fCellVoltage := 0.0;        // 复核失败回缺省 / Fallback on recheck failure
    fOhmicDrop := 0.0;          // 复核失败回缺省 / Fallback on recheck failure
    uErrorId := 16#0002_9214;   // 出口非有限拒收 / Output non-finite reject
    RETURN;
END_IF
IF (fCellVoltage < 2.0) OR (fCellVoltage > 8.0) THEN
    uErrorId := 16#0002_9214;   // 信息级：槽电压出工艺窗 / Info: voltage out of window
    RETURN;                     // bValid 保持 FALSE / Validity stays false
END_IF
bValid := TRUE;                 // 有效回执 / Validity receipt
FC_DL_PotlineCellVoltageBudgetCalc := fCellVoltage;     // 返回值镜像槽电压 / Return mirrors voltage
END_FUNCTION

(* ---- FC_DL_PotlineCrustBreakerEnergyCalc.st ---- *)
// FC_DL_PotlineCrustBreakerEnergyCalc v1.0.0
// 开源溯源：clean-room 自研（族 DL_Process，ST 生态实测 0 命中，无外部代码引入）
(*
  功能: 打壳机械能：单次冲击 = F[kN]·s[mm]/1000 [kJ]（kN·mm = J，除 1000 得 kJ），
        单次打壳 = 单次冲击 × 冲击数，平均功率 = 单次打壳 × 频次/3600 [kW]（kJ/h ÷ 3600 = kW）。
  邻件/码位: 与 FC_DL_PotlineAnodeEffectEnergyCalc 同为能耗件（本件机械能 vs 电能，不可互换）；
             16#0002_9219 = 非有限、任一量非正或冲击数 < 1 拒收。
*)
FUNCTION FC_DL_PotlineCrustBreakerEnergyCalc : REAL
VAR_INPUT
    fImpactForce     : REAL := 20.0;   // 单次冲击力 [kN]，域 > 0 / Impact force [kN]
    fStroke          : REAL := 50.0;   // 冲击行程 [mm]，域 > 0 / Impact stroke [mm]
    fStrikesPerBreak : REAL := 3.0;    // 单次打壳冲击数 [次]，域 >= 1 / Strikes per break [count]
    fBreaksPerHour   : REAL := 6.0;    // 打壳频次 [次/h]，域 > 0 / Breaks per hour [count/h]
END_VAR
VAR_OUTPUT
    fEnergyPerBreak : REAL;             // 单次打壳机械能 [kJ] / Energy per break [kJ]
    fPowerAvg       : REAL;             // 平均功率 [kW] / Average mechanical power [kW]
    bValid          : BOOL;             // 结果有效回执 [-] / Result validity receipt
    uErrorId        : UDINT;            // 事件码，0 = 无事件 / Event code
END_VAR
VAR
    fEnergyPerStrike : REAL := 0.0;     // 单次冲击机械能 [kJ] / Energy per strike [kJ]
END_VAR
// 段 0：全路径出口安全缺省 / Safe defaults on all outlets
fEnergyPerBreak := 0.0;                 // 单次打壳能量缺省零 / Per-break energy default zero
fPowerAvg := 0.0;                       // 平均功率缺省零 / Average power default zero
bValid := FALSE;                        // 有效回执预清 / Validity preset clear
uErrorId := 16#0000;                    // 事件码预清 / Event code preset clear
FC_DL_PotlineCrustBreakerEnergyCalc := 0.0; // 返回值缺省零（镜像单次能量）/ Return default zero
// 段 1：非有限闸（四入参全枚举）/ Non-finite gate over all inputs
IF (fImpactForce <> fImpactForce) OR (fStroke <> fStroke)
   OR (fStrikesPerBreak <> fStrikesPerBreak) OR (fBreaksPerHour <> fBreaksPerHour)
   OR (ABS(fImpactForce) >= 3.0E38) OR (ABS(fStroke) >= 3.0E38)
   OR (ABS(fStrikesPerBreak) >= 3.0E38) OR (ABS(fBreaksPerHour) >= 3.0E38) THEN
    uErrorId := 16#0002_9219;   // 入参非有限拒收 / Non-finite input reject
    RETURN;
END_IF
// 段 2：域闸（力/行程/频次为正 + 冲击数下限，R4）/ Domain gate
IF (fImpactForce <= 0.0) OR (fStroke <= 0.0) OR (fBreaksPerHour <= 0.0) THEN
    uErrorId := 16#0002_9219;   // 力、行程或频次非正 / Non-positive force, stroke or rate
    RETURN;
END_IF
IF fStrikesPerBreak < 1.0 THEN
    uErrorId := 16#0002_9219;   // 冲击数不足 1 次 / Strike count below one
    RETURN;
END_IF
// 段 3：主计算（冲击能 → 单次打壳能 → 平均功率）/ Main computation
fEnergyPerStrike := fImpactForce * fStroke / 1000.0;            // F·s/1000 [kJ] / Energy per strike
fEnergyPerBreak := fEnergyPerStrike * fStrikesPerBreak;         // 单次打壳机械能 [kJ] / Per break
fPowerAvg := fEnergyPerBreak * fBreaksPerHour / 3600.0;         // 平均功率 [kW] / Average power
// 段 4：出口闸（双输出非有限复核 + 非负复核）/ Outlet gate
IF (fEnergyPerBreak <> fEnergyPerBreak) OR (fPowerAvg <> fPowerAvg)
   OR (ABS(fEnergyPerBreak) >= 3.0E38) OR (ABS(fPowerAvg) >= 3.0E38)
   OR (fEnergyPerBreak < 0.0) OR (fPowerAvg < 0.0) THEN
    fEnergyPerBreak := 0.0;     // 复核失败回缺省 / Fallback on recheck failure
    fPowerAvg := 0.0;           // 复核失败回缺省 / Fallback on recheck failure
    uErrorId := 16#0002_9219;   // 出口复核拒收 / Output recheck reject
    RETURN;
END_IF
bValid := TRUE;                 // 有效回执 / Validity receipt
FC_DL_PotlineCrustBreakerEnergyCalc := fEnergyPerBreak;     // 返回值镜像单次机械能 / Return mirrors
END_FUNCTION

(* ---- FC_DL_PotlineCurrentEfficiencyCalc.st ---- *)
// FC_DL_PotlineCurrentEfficiencyCalc v1.0.0
// 开源溯源：clean-room 自研（族 DL_Process，ST 生态实测 0 命中，无外部代码引入）
(*
  功能: 电流效率反算：理论产铝 = I[kA]·0.3355·t[h] [kg]，CE = 100·实测/理论 [%]；
        CE > 105% 判计量异常（产物称重或电流计量故障）。
  邻件/码位: 与 FC_DL_PotlineAluminaFeedRateCalc 互为逆过程（本件由实测反推 CE）；
             16#0002_9215 = 非有限、理论量近零或 CE 越 105% 上限。
*)
FUNCTION FC_DL_PotlineCurrentEfficiencyCalc : REAL
VAR_INPUT
    fActualAlKg : REAL := 1000.0;   // 统计期内实测产铝 [kg]，域 >= 0 / Measured mass [kg]
    fCurrentKA  : REAL := 400.0;    // 系列电流 [kA]，域 > 0 / Line current [kA]
    fHours      : REAL := 24.0;     // 统计时长 [h]，域 > 0 / Statistics window [h]
END_VAR
VAR_OUTPUT
    fCE      : REAL;                // 电流效率 [%] / Current efficiency [%]
    bValid   : BOOL;                // 结果有效回执 [-] / Result validity receipt
    uErrorId : UDINT;               // 事件码，0 = 无事件 / Event code
END_VAR
VAR
    fTheory : REAL := 0.0;          // 理论产铝量 [kg] / Theoretical mass [kg]
END_VAR
// 段 0：全路径出口安全缺省 / Safe defaults on all outlets
fCE := 0.0;                     // 电流效率缺省零 / Current efficiency default zero
bValid := FALSE;                // 有效回执预清 / Validity preset clear
uErrorId := 16#0000;            // 事件码预清 / Event code preset clear
FC_DL_PotlineCurrentEfficiencyCalc := 0.0;  // 返回值缺省零（镜像 CE）/ Return default zero
// 段 1：非有限闸（三入参全枚举）/ Non-finite gate over all inputs
IF (fActualAlKg <> fActualAlKg) OR (fCurrentKA <> fCurrentKA) OR (fHours <> fHours)
   OR (ABS(fActualAlKg) >= 3.0E38) OR (ABS(fCurrentKA) >= 3.0E38) OR (ABS(fHours) >= 3.0E38) THEN
    uErrorId := 16#0002_9215;   // 入参非有限拒收 / Non-finite input reject
    RETURN;
END_IF
// 段 2：域闸（实测非负 + 电流与时长为正防除零，R4）/ Domain gate
IF fActualAlKg < 0.0 THEN
    uErrorId := 16#0002_9215;   // 实测产铝为负 / Negative measured mass
    RETURN;
END_IF
IF (fCurrentKA <= 1.0E-6) OR (fHours <= 1.0E-6) THEN
    uErrorId := 16#0002_9215;   // 电流或时长非正 / Non-positive current or window
    RETURN;
END_IF
// 段 3：主计算（理论量 → CE）/ Main computation
fTheory := fCurrentKA * 0.3355 * fHours;                        // 理论产铝量 / Theoretical mass
IF fTheory <= 1.0E-6 THEN
    uErrorId := 16#0002_9215;   // 理论量近零，CE 不可解 / Theoretical mass too small
    RETURN;
END_IF
fCE := 100.0 * fActualAlKg / fTheory;                           // CE = 100·实测/理论 / Efficiency
// 段 4：出口闸（非有限复核 + 105% 计量异常判定）/ Outlet gate
IF (fCE <> fCE) OR (ABS(fCE) >= 3.0E38) THEN
    fCE := 0.0;                 // 复核失败回缺省 / Fallback on recheck failure
    uErrorId := 16#0002_9215;   // 出口非有限拒收 / Output non-finite reject
    RETURN;
END_IF
IF fCE > 105.0 THEN
    uErrorId := 16#0002_9215;   // 信息级：CE 超 105% 判计量异常 / Info: metrology anomaly
    RETURN;                     // bValid 保持 FALSE / Validity stays false
END_IF
bValid := TRUE;                 // 有效回执 / Validity receipt
FC_DL_PotlineCurrentEfficiencyCalc := fCE;      // 返回值镜像 CE / Return mirrors efficiency
END_FUNCTION

(* ---- FC_DL_PotlineMetalLevelCalc.st ---- *)
// FC_DL_PotlineMetalLevelCalc v1.0.0
// 开源溯源：clean-room 自研（族 DL_Process，ST 生态实测 0 命中，无外部代码引入）
(*
  功能: 铝水平 = m/(ρ·A)·100 [cm]（m³/m² = m，再 ×100 转 cm），电解质水平 = 铝水平 + 电解质层厚；
        密度入参为 1.0（占位缺省，调用方未组态）时改用 2300.0 kg/m³。
  邻件/码位: 与 FC_DL_PotlineBathTempDeviationCalc 同族不同域（几何液位 vs 热状态）；
             16#0002_9217 = 非有限、面积或密度非正、层厚为负拒收。
*)
FUNCTION FC_DL_PotlineMetalLevelCalc : REAL
VAR_INPUT
    fMetalMassKg  : REAL := 10000.0;    // 槽内铝量 [kg]，域 >= 0 / Metal mass in cell [kg]
    fCavityArea   : REAL := 25.0;       // 槽膛面积 [m²]，域 > 0 / Cavity area [m^2]
    fBathDepth    : REAL := 20.0;       // 电解质层厚 [cm]，域 >= 0 / Bath layer depth [cm]
    fMetalDensity : REAL := 2300.0;     // 铝液密度 [kg/m³]，域 > 0 / Metal density [kg/m^3]
END_VAR
VAR_OUTPUT
    fMetalLevel : REAL;                 // 铝水平 [cm] / Metal level [cm]
    fBathLevel  : REAL;                 // 电解质水平 [cm] / Bath level [cm]
    bValid      : BOOL;                 // 结果有效回执 [-] / Result validity receipt
    uErrorId    : UDINT;                // 事件码，0 = 无事件 / Event code
END_VAR
VAR
    fDensity : REAL := 0.0;             // 生效密度 [kg/m³] / Effective density [kg/m^3]
END_VAR
// 段 0：全路径出口安全缺省 / Safe defaults on all outlets
fMetalLevel := 0.0;                 // 铝水平缺省零 / Metal level default zero
fBathLevel := 0.0;                  // 电解质水平缺省零 / Bath level default zero
bValid := FALSE;                    // 有效回执预清 / Validity preset clear
uErrorId := 16#0000;                // 事件码预清 / Event code preset clear
FC_DL_PotlineMetalLevelCalc := 0.0;         // 返回值缺省零（镜像铝水平）/ Return default zero
// 段 1：非有限闸（四入参全枚举）/ Non-finite gate over all inputs
IF (fMetalMassKg <> fMetalMassKg) OR (fCavityArea <> fCavityArea)
   OR (fBathDepth <> fBathDepth) OR (fMetalDensity <> fMetalDensity)
   OR (ABS(fMetalMassKg) >= 3.0E38) OR (ABS(fCavityArea) >= 3.0E38)
   OR (ABS(fBathDepth) >= 3.0E38) OR (ABS(fMetalDensity) >= 3.0E38) THEN
    uErrorId := 16#0002_9217;   // 入参非有限拒收 / Non-finite input reject
    RETURN;
END_IF
// 段 2：域闸（面积与密度为正 + 层厚非负 + 密度占位替换，R4）/ Domain gate
IF (fCavityArea <= 1.0E-6) OR (fMetalDensity <= 0.0) THEN
    uErrorId := 16#0002_9217;   // 面积或密度非正，液位不可解 / Non-positive area or density
    RETURN;
END_IF
IF fBathDepth < 0.0 THEN
    uErrorId := 16#0002_9217;   // 电解质层厚为负 / Negative bath depth
    RETURN;
END_IF
fDensity := fMetalDensity;                                      // 密度先直取 / Take density as-is
IF fDensity <= 1.0 THEN
    fDensity := 2300.0;                                         // 占位缺省替换 / Placeholder replaced
END_IF
// 段 3：主计算（质量→体积→液位）/ Main computation
fMetalLevel := fMetalMassKg / (fDensity * fCavityArea) * 100.0;     // 铝水平 [cm] / Metal level
fBathLevel := fMetalLevel + fBathDepth;                             // 电解质水平 [cm] / Bath level
// 段 4：出口闸（双输出非有限复核 + 非负复核）/ Outlet gate
IF (fMetalLevel <> fMetalLevel) OR (fBathLevel <> fBathLevel)
   OR (ABS(fMetalLevel) >= 3.0E38) OR (ABS(fBathLevel) >= 3.0E38)
   OR (fMetalLevel < 0.0) OR (fBathLevel < 0.0) THEN
    fMetalLevel := 0.0;         // 复核失败回缺省 / Fallback on recheck failure
    fBathLevel := 0.0;          // 复核失败回缺省 / Fallback on recheck failure
    uErrorId := 16#0002_9217;   // 出口复核拒收 / Output recheck reject
    RETURN;
END_IF
bValid := TRUE;                 // 有效回执 / Validity receipt
FC_DL_PotlineMetalLevelCalc := fMetalLevel;     // 返回值镜像铝水平 / Return mirrors metal level
END_FUNCTION

(* ---- FC_DL_PouringTimeCalc.st ---- *)
(*
 * FC_DL_PouringTimeCalc | C2 | DL_Process
 * 功能：浇注时间估算（浇注重量平方根经验式）与上下限钳位       单位：重量 [kg]、系数 [s/√kg]、时间 [s]
 * 工况边界：经验式 t = k×√G，k 取 1.8 s/√kg（灰铸铁中小件典型值）；仅适用于重力浇注且浇口未更换的场合；重量须 >0、系数须 >0 且有限；超出 [min,max] 时钳位并置 xClamped（判据取自未钳位原值，R24）
 * 代数值回代：G=50 kg、k=1.8 → t=1.8×7.071=12.73 s，落在 [4,30] → xClamped=FALSE（与 spec 回代行一致）
 * 开源溯源：clean-room 自研，未复制任何第三方代码（无外部来源）
 *)
FUNCTION FC_DL_PouringTimeCalc : BOOL
VAR_INPUT
    rPourWeightKg : REAL := 50.0;     // 浇注重量（含浇冒口）| pouring weight including gating and risers [kg]
    rCoeff        : REAL := 1.8;      // 经验系数 | empirical coefficient [s/√kg]
    rMinS         : REAL := 4.0;      // 允许最短浇注时间 | minimum pouring time [s]
    rMaxS         : REAL := 30.0;     // 允许最长浇注时间 | maximum pouring time [s]
END_VAR
VAR_OUTPUT
    rPourTimeS : REAL;                // 浇注时间设定 | pouring time setpoint [s]
    rRawTimeS  : REAL;                // 未钳位的原始计算值 | raw time before clamping [s]
    xClamped   : BOOL;                // 已打限幅（信息级）| clamped against the limits, informational
    xValid     : BOOL;                // 输出有效 | outputs valid
END_VAR
VAR
    xFinG  : BOOL;                    // 重量有限性 | weight is finite
    xFinK  : BOOL;                    // 系数有限性 | coefficient is finite
    xFinLo : BOOL;                    // 下限有限性 | lower limit is finite
    xFinHi : BOOL;                    // 上限有限性 | upper limit is finite
END_VAR
VAR CONSTANT
    DL_PTC_EPS : REAL := 1.0E-6;      // 浮点比较容差 | floating comparison tolerance [s]
END_VAR

// 段1｜非有限闸（R19）
xFinG := (rPourWeightKg = rPourWeightKg) AND ((rPourWeightKg - rPourWeightKg) = 0.0);
xFinK := (rCoeff = rCoeff) AND ((rCoeff - rCoeff) = 0.0);
xFinLo := (rMinS = rMinS) AND ((rMinS - rMinS) = 0.0);
xFinHi := (rMaxS = rMaxS) AND ((rMaxS - rMaxS) = 0.0);
IF (NOT xFinG) OR (NOT xFinK) OR (NOT xFinLo) OR (NOT xFinHi) THEN
    rPourTimeS := 4.0;                // 安全值：取下限（快速浇注侧不可取，取允许最短）| safe value, the shortest permitted time
    rRawTimeS := 4.0;
    xClamped := TRUE;
    xValid := FALSE;
    FC_DL_PouringTimeCalc := FALSE;
    RETURN;
END_IF

// 段2｜域闸：重量与系数须为正（√G 的定义域），限幅区间须有效
IF (rPourWeightKg <= 0.0) OR (rCoeff <= 0.0) OR (rMaxS <= rMinS) THEN
    rPourTimeS := rMinS;              // 安全值：取下限 | safe value, the lower limit
    rRawTimeS := rMinS;
    xClamped := TRUE;
    xValid := FALSE;
    FC_DL_PouringTimeCalc := FALSE;
    RETURN;
END_IF

// 段3｜算法：t = k×√G
rRawTimeS := rCoeff * SQRT(rPourWeightKg);

// 段4｜限幅与打限标志（判据取自未钳位原值，R24）
xClamped := (rRawTimeS > (rMaxS + DL_PTC_EPS)) OR (rRawTimeS < (rMinS - DL_PTC_EPS));
rPourTimeS := LIMIT(rMinS, rRawTimeS, rMaxS);

// 段5｜出口
xValid := TRUE;
FC_DL_PouringTimeCalc := TRUE;
END_FUNCTION

(* ---- FC_DL_PowderFillDensityCalc.st ---- *)
(*
  Component : FC_DL_PowderFillDensityCalc
  Category  : DL_Process
  Type      : FC
  Complexity: C1
  VERSION   : v1.0.0
  功能      : 装粉松装密度与填充高度核算：按粉重、模腔面积与松装密度算填充容积与填充高度，并给出压制压缩比。
  开源溯源  : 道莅原创 clean-room 自研（无外部代码引用）｜License: MIT
  边界条件  : ① 模腔面积与松装密度须 > 1e-9，否则返回哨兵 -1（松装密度为除子）；
              ② 压缩比为压坯密度与松装密度之比，压坯密度为 0 时回 1.0（无压缩）；
              ③ 量纲链：kg→g 除 g/cm³ 得 cm³，再乘 1000 除 mm² 得 mm。
*)
FUNCTION FC_DL_PowderFillDensityCalc : REAL
VAR_INPUT
    fPowderKg     : REAL;   (* 单件装粉质量 [kg] Powder mass per part *)
    fCavityAreaMm2: REAL;   (* 模腔投影面积 [mm²] Cavity cross-section area *)
    fAppDensGcm3  : REAL;   (* 粉末松装密度 [g/cm³] Apparent density *)
    fPressDensGcm3: REAL;   (* 压坯密度 [g/cm³] Green compact density *)
END_VAR
VAR_OUTPUT
    fFillVolCm3 : REAL;   (* 填充容积 [cm³] Fill volume *)
    fFillHeightMm: REAL;  (* 填充高度 [mm] Fill height *)
    fCompRatio  : REAL;   (* 压缩比（压坯/松装） [-] Compression ratio *)
    xValid      : BOOL;   (* 计算有效性标志 [-] Calculation valid flag *)
END_VAR
VAR CONSTANT
    DL_EPS       : REAL := 1.0E-9;   (* 除零判定容差 [无量纲] Divide-by-zero tolerance *)
    DL_G_PER_KG  : REAL := 1000.0;   (* 千克转克系数 [g/kg] Grams per kilogram *)
    DL_MM3_PER_CM3: REAL := 1000.0;  (* 立方厘米转立方毫米 [mm³/cm³] mm3 per cm3 *)
    DL_ZERO      : REAL := 0.0;      (* 零常量 [无量纲] Zero constant *)
END_VAR
(* 出口预置：四出口统一预置 *)
fFillVolCm3 := 0.0; fFillHeightMm := 0.0; fCompRatio := 1.0; xValid := FALSE;
(* 非有限拦截：自反判 NaN，自身差值判 Inf *)
IF (fPowderKg <> fPowderKg) OR ((fPowderKg - fPowderKg) <> 0.0)
   OR (fCavityAreaMm2 <> fCavityAreaMm2) OR ((fCavityAreaMm2 - fCavityAreaMm2) <> 0.0)
   OR (fAppDensGcm3 <> fAppDensGcm3) OR ((fAppDensGcm3 - fAppDensGcm3) <> 0.0)
   OR (fPressDensGcm3 <> fPressDensGcm3) OR ((fPressDensGcm3 - fPressDensGcm3) <> 0.0) THEN
    FC_DL_PowderFillDensityCalc := -1.0;  (* 哨兵 -1：输入非有限 / Sentinel -1 non-finite *)
    RETURN;
END_IF
(* 组态域闸：面积与松装密度均为除子，粉重须非负 *)
IF (fCavityAreaMm2 <= DL_EPS) OR (fAppDensGcm3 <= DL_EPS) OR (fPowderKg < DL_ZERO) THEN
    FC_DL_PowderFillDensityCalc := -1.0;  (* 哨兵 -1：组态非法 / Sentinel -1 bad config *)
    RETURN;
END_IF
(* 填充容积：V = m / 松装密度 [cm³]，分母已过域闸 *)
fFillVolCm3 := (fPowderKg * DL_G_PER_KG) / fAppDensGcm3;
(* 填充高度：h = V(mm³) / A(mm²) [mm] *)
fFillHeightMm := (fFillVolCm3 * DL_MM3_PER_CM3) / fCavityAreaMm2;
(* 压缩比：压坯密度 / 松装密度，压坯密度为 0 时保持 1.0 *)
IF fPressDensGcm3 > DL_EPS THEN
    fCompRatio := fPressDensGcm3 / fAppDensGcm3;
ELSE
    fCompRatio := 1.0;                    (* 无压坯数据：按无压缩处理 *)
END_IF
xValid := TRUE;                           (* 链路有效 / Chain valid *)
FC_DL_PowderFillDensityCalc := fFillHeightMm;  (* 返回填充高度 [mm] / Return fill height *)
END_FUNCTION

(* ---- FC_DL_PreheaterCyclonePressureCalc.st ---- *)
(*
  Name: FC_DL_PreheaterCyclonePressureCalc
  Category: DL_Process
  Version: 1.0.0
  Round: R91 / 2026-11-25
  开源溯源：clean-room 自研（族 水泥窑篦冷机与预热器，ST 开源生态实测 0 命中，无外部代码引入）
  功能：1) 旋风筒压损按局部阻力式 dP = zeta * rho * v^2 / 2 计算，再折 kPa：
           fCycloneDpKpa = zeta * fGasDensityKgm3 * v^2 / 2 / 1000，
           其中 zeta 为旋风筒进出口综合阻力系数（含内筒插入深度经验项）。
        2) 负荷率 fDpLoadPct = 压损 / 设备许可压损上限 * 100，用于判断系统是否接近风机能力极限。
        3) 堵塞风险判据：入口风速低于 fVelBlockMs 时判 xBlockRisk（低风速不能维持旋流的
           携带能力，粉尘易在锥体沉积），该判据与压损超限判据并行独立输出。
  边界条件：1) 非有限值闸：五路实值入参先过 NOT(x > -DL_BIG AND x < DL_BIG)，同时拦 NaN 与 Inf，
           命中即闸断实值通路（全部输出强制 0.0），不得只置标志（R19）。
        2) 分母零闸：设备许可压损上限 fDpMaxKpa 必须 > DL_EPS（负荷率的分母），否则判无效。
        3) 物理域闸：气体密度 fGasDensityKgm3 必须 > 0（密度为零即非真实气体），
           阻力系数 fResistCoef 必须 > 0，入口风速不得为负；任一越界判无效，不钳制。
        4) 风速上限：入口风速超过 DL_VEL_HI_MS 判无效（超上限说明测点或管径组态错误，
           此时压损式的外推已失真），不把超限值当作高风速使用。
        5) 判据取原始值（R24）：压损越限判定使用钳制前的 _fDpRawKpa。
        6) 物理域钳制：压损钳 0.0 ~ fDpMaxKpa；负荷率钳 0.0 ~ DL_PCT_HI；风速只判不钳（供观测）。
  量纲自证：zeta 无因次；rho*v^2/2 = (kg/m3)*(m2/s2) = kg/(m*s2) = Pa；
           除以 1000 得 kPa，故 fCycloneDpKpa 量纲为 [kPa]；
           fDpLoadPct = (kPa)/(kPa)*100 = 无因次百分数 [%]，量纲合法。
  修订历史 Revision :
    2026-11-25  v1.0.0  R91 首版
*)

FUNCTION FC_DL_PreheaterCyclonePressureCalc : BOOL
VAR_INPUT
    fInletVelMs      : REAL;   // 旋风筒入口风速 [m/s] / Cyclone inlet gas velocity [m/s]
    fResistCoef      : REAL;   // 综合阻力系数（无因次）[-] / Combined resistance coefficient [-]
    fGasDensityKgm3  : REAL;   // 工况气体密度 [kg/m3] / Gas density at working condition [kg/m3]
    fDpMaxKpa        : REAL;   // 设备许可压损上限 [kPa] / Permitted pressure drop [kPa]
    fVelBlockMs      : REAL;   // 堵塞风险风速下限 [m/s] / Blockage-risk velocity low limit [m/s]
END_VAR
VAR_OUTPUT
    fCycloneDpKpa    : REAL;   // 旋风筒压损 [kPa] / Cyclone pressure drop [kPa]
    fDpLoadPct       : REAL;   // 压损负荷率 [%] / Pressure drop load ratio [%]
    xDpOver          : BOOL;   // 压损超限标志 [bool] / Pressure drop overrun flag [bool]
    xBlockRisk       : BOOL;   // 堵塞风险标志（入口风速不足）[bool] / Blockage risk flag [bool]
    xValid           : BOOL;   // 计算有效标志 [bool] / Calculation valid flag [bool]
END_VAR
VAR
    _fDynPa          : REAL;   // 动压 [Pa] / Dynamic pressure [Pa]
    _fDpRawKpa       : REAL;   // 钳制前的原始压损 [kPa] / Raw pressure drop before limiting [kPa]
    _fLoadRawPct     : REAL;   // 钳制前的原始负荷率 [%] / Raw load ratio before limiting [%]
END_VAR
VAR CONSTANT
    DL_EPS           : REAL := 1.0E-9;    // 数值零闸阈值 [-] / Numeric zero gate threshold [-]
    DL_BIG           : REAL := 1.0E12;    // 非有限值闸量级上限 [-] / Finiteness gate magnitude [-]
    DL_TWO           : REAL := 2.0;       // 动压式系数分母（v^2/2）[-] / Dynamic pressure divisor [-]
    DL_PA_PER_KPA    : REAL := 1000.0;    // 帕到千帕的折算 [Pa/kPa] / Pascals per kilopascal [Pa/kPa]
    DL_PCT           : REAL := 100.0;     // 百分比换算因子 [%] / Percent conversion factor [%]
    DL_PCT_HI        : REAL := 100.0;     // 负荷率物理上限 [%] / Load ratio upper bound [%]
    DL_VEL_HI_MS     : REAL := 40.0;      // 入口风速组态上限 [m/s] / Inlet velocity configuration upper bound [m/s]
END_VAR

(* —— 段 1：非有限值闸（R19：闸断实值通路） —— *)
IF NOT (fInletVelMs > -DL_BIG AND fInletVelMs < DL_BIG)
   OR NOT (fResistCoef > -DL_BIG AND fResistCoef < DL_BIG)
   OR NOT (fGasDensityKgm3 > -DL_BIG AND fGasDensityKgm3 < DL_BIG)
   OR NOT (fDpMaxKpa > -DL_BIG AND fDpMaxKpa < DL_BIG)
   OR NOT (fVelBlockMs > -DL_BIG AND fVelBlockMs < DL_BIG) THEN
    fCycloneDpKpa := 0.0;                   // 输出强制 0.0，切断污染源 / Force zero, cut polluted path
    fDpLoadPct := 0.0;                      // 负荷率强制 0.0 / Load ratio forced to zero
    xDpOver := FALSE;                       // 失效侧超限位保持假 / Overrun stays false
    xBlockRisk := FALSE;                    // 失效侧堵塞风险位保持假 / Blockage risk stays false
    xValid := FALSE;                        // 有效位清零 / Validity cleared
    FC_DL_PreheaterCyclonePressureCalc := FALSE;   // 返回码与有效位同源 / Return mirrors validity
    RETURN;                                 // 立即退出 / Immediate exit
END_IF

(* —— 段 2：分母零闸与物理域闸（负荷率分母 + 密度/系数必须为正） —— *)
IF (fDpMaxKpa <= DL_EPS)                                          // 压损上限必须已组态
   OR (fGasDensityKgm3 <= DL_EPS)                                 // 气体密度必须为正
   OR (fResistCoef <= DL_EPS)                                     // 阻力系数必须为正
   OR (fInletVelMs < 0.0)                                         // 风速不得为负
   OR (fVelBlockMs < 0.0)                                         // 堵塞下限不得为负
   OR (fInletVelMs > DL_VEL_HI_MS) THEN                           // 风速超组态上限：测点或管径错误
    fCycloneDpKpa := 0.0;                   // 参数不可用即无压损 / No parameter, no pressure drop
    fDpLoadPct := 0.0;                      // 负荷率不可算 / Load ratio not computable
    xDpOver := FALSE;                       // 失效侧超限位保持假 / Overrun stays false
    xBlockRisk := FALSE;                    // 失效侧堵塞风险位保持假 / Blockage risk stays false
    xValid := FALSE;                        // 判无效 / Invalid
    FC_DL_PreheaterCyclonePressureCalc := FALSE;   // 返回码同步 / Return synchronised
    RETURN;                                 // 提前退出 / Early exit
END_IF

(* —— 段 3：主算式（不钳制，先出原始值供段 4 判据使用，R24） —— *)
_fDynPa := fGasDensityKgm3 * fInletVelMs * fInletVelMs / DL_TWO;                  // 动压 [Pa]
_fDpRawKpa := fResistCoef * _fDynPa / DL_PA_PER_KPA;                              // 压损 [kPa]
_fLoadRawPct := _fDpRawKpa / fDpMaxKpa * DL_PCT;                                  // 负荷率 [%]

(* —— 段 4：判据（取原始值；单点 BOOL 聚合避免多处赋 FALSE 覆盖） —— *)
xDpOver := (_fDpRawKpa > fDpMaxKpa);                                              // 压损越许可上限
xBlockRisk := (fInletVelMs < fVelBlockMs);                                        // 风速不足：旋流携带能力丧失
xValid := (fVelBlockMs < DL_VEL_HI_MS)                                            // 堵塞下限须低于组态上限（否则判据恒真）
          AND (_fLoadRawPct >= 0.0);                                              // 负荷率不得为负

(* —— 段 5：输出单点写盘（钳制到物理域内，判定结果已在段 4 定案） —— *)
fCycloneDpKpa := LIMIT(0.0, _fDpRawKpa, fDpMaxKpa);                               // 压损钳 0..上限 [kPa]
fDpLoadPct := LIMIT(0.0, _fLoadRawPct, DL_PCT_HI);                                // 负荷率钳 0..100 [%]
FC_DL_PreheaterCyclonePressureCalc := xValid;                                     // 返回码：TRUE = 计算可信

END_FUNCTION

(* ---- FC_DL_PreheaterStageEfficiencyCalc.st ---- *)
(*
  Name: FC_DL_PreheaterStageEfficiencyCalc
  Category: DL_Process
  Version: 1.0.0
  Round: R91 / 2026-11-25
  开源溯源：clean-room 自研（族 水泥窑篦冷机与预热器，ST 开源生态实测 0 命中，无外部代码引入）
  功能：1) 预热器单级换热效率按「气体放热占理论最大放热的比例」计算：
           eff = (T_gasIn − T_gasOut) / (T_gasIn − T_matIn) * 100，
           分母是气体入口温度与物料入口温度之差，即可传给物料的温度势上限；
           方向固定不可交换（气体为热源、物料为受热体）。
        2) 派生输出：气体温降 fGasDropK 与出口逼近温差 fApproachK = T_gasOut − T_matIn，
           后者是级间结皮/堵塞的早期征兆量（逼近温差过小意味着换热面积不足或物料短路）。
        3) 效率物理域校验：效率必须落在 0.0 ~ 100.0 % 且不超过该级设计上限 fEffMaxPct；
           超上限在热力学上不可能，判为温度测点故障而非换热优异。
  边界条件：1) 非有限值闸：四路实值入参先过 NOT(x > -DL_BIG AND x < DL_BIG)，同时拦 NaN 与 Inf，
           命中即闸断实值通路（全部输出强制 0.0），不得只置标志（R19）。
        2) 分母零闸：温度势 |T_gasIn − T_matIn| <= DL_EPS 时不做除法（进出口等温即无势差），
           全部输出清零并判无效。
        3) 温度势方向闸：T_gasIn 必须严格高于 T_matIn，否则热流反向（物料比气体还热），判无效。
        4) 设计上限域闸：fEffMaxPct 必须落在 (0.0, 100.0] 内，越域视为未组态判无效，不做钳制。
        5) 判据取原始值（R24）：效率越限判定使用钳制前的 _fEffRawPct，不得先钳再判。
        6) 物理域钳制：效率钳 0.0 ~ 100.0 %；温降与逼近温差钳 >= 0（负值属测点反向，另由 xValid 拦截）。
  量纲自证：fGasDropK = (degC) − (degC) = (K)；fApproachK = (degC) − (degC) = (K)；
           fEffPct = (K)/(K)*100 = 无因次百分数 [%]，比量两侧同为温差量纲，量纲关系合法。
  修订历史 Revision :
    2026-11-25  v1.0.0  R91 首版
*)

FUNCTION FC_DL_PreheaterStageEfficiencyCalc : BOOL
VAR_INPUT
    fGasInC          : REAL;   // 该级进口气体温度 [degC] / Stage inlet gas temperature [degC]
    fGasOutC         : REAL;   // 该级出口气体温度 [degC] / Stage outlet gas temperature [degC]
    fMatInC          : REAL;   // 该级进口物料温度 [degC] / Stage inlet material temperature [degC]
    fEffMaxPct       : REAL;   // 该级设计换热效率上限 [%] / Design efficiency upper limit [%]
END_VAR
VAR_OUTPUT
    fEffPct          : REAL;   // 单级换热效率 [%] / Single-stage heat exchange efficiency [%]
    fGasDropK        : REAL;   // 气体温降 [K] / Gas temperature drop [K]
    fApproachK       : REAL;   // 出口气体与进口物料的逼近温差 [K] / Outlet approach temperature [K]
    xEffOver         : BOOL;   // 效率超设计上限标志 [bool] / Efficiency over design limit flag [bool]
    xValid           : BOOL;   // 计算有效标志 [bool] / Calculation valid flag [bool]
END_VAR
VAR
    _fPotentialK     : REAL;   // 温度势（气体入口 − 物料入口）[K] / Temperature potential [K]
    _fDropRawK       : REAL;   // 钳制前的气体温降 [K] / Raw gas temperature drop [K]
    _fApproachRawK   : REAL;   // 钳制前的逼近温差 [K] / Raw approach temperature [K]
    _fEffRawPct      : REAL;   // 钳制前的原始效率 [%] / Raw efficiency before limiting [%]
END_VAR
VAR CONSTANT
    DL_EPS           : REAL := 1.0E-9;    // 数值零闸阈值 [-] / Numeric zero gate threshold [-]
    DL_BIG           : REAL := 1.0E12;    // 非有限值闸量级上限 [-] / Finiteness gate magnitude [-]
    DL_PCT           : REAL := 100.0;     // 百分比换算因子 [%] / Percent conversion factor [%]
    DL_EFF_LO_PCT    : REAL := 0.0;       // 效率物理域下限 [%] / Efficiency physical domain low [%]
    DL_EFF_HI_PCT    : REAL := 100.0;     // 效率物理域上限 [%] / Efficiency physical domain high [%]
    DL_ZERO_K        : REAL := 0.0;       // 温差零基准 [K] / Zero temperature-difference reference [K]
END_VAR

(* —— 段 1：非有限值闸（R19：闸断实值通路） —— *)
IF NOT (fGasInC > -DL_BIG AND fGasInC < DL_BIG)
   OR NOT (fGasOutC > -DL_BIG AND fGasOutC < DL_BIG)
   OR NOT (fMatInC > -DL_BIG AND fMatInC < DL_BIG)
   OR NOT (fEffMaxPct > -DL_BIG AND fEffMaxPct < DL_BIG) THEN
    fEffPct := 0.0;                         // 输出强制 0.0，切断污染源 / Force zero, cut polluted path
    fGasDropK := 0.0;                       // 温降强制 0.0 / Gas drop forced to zero
    fApproachK := 0.0;                      // 逼近温差强制 0.0 / Approach forced to zero
    xEffOver := FALSE;                      // 失效侧超限位保持假 / Overrun stays false when invalid
    xValid := FALSE;                        // 有效位清零 / Validity cleared
    FC_DL_PreheaterStageEfficiencyCalc := FALSE;   // 返回码与有效位同源 / Return mirrors validity
    RETURN;                                 // 立即退出 / Immediate exit
END_IF

(* —— 段 2：温度势方向闸与分母零闸（分母为温度势，必须先验方向再验量级） —— *)
_fPotentialK := fGasInC - fMatInC;                                                // 温度势 [K]
IF (_fPotentialK <= DL_EPS) THEN                                                  // 势差为零或反向：无换热驱动力
    fEffPct := 0.0;                         // 无势差即无效率 / No potential, no efficiency
    fGasDropK := 0.0;                       // 温降不可算 / Drop not computable
    fApproachK := 0.0;                      // 逼近温差不可算 / Approach not computable
    xEffOver := FALSE;                      // 失效侧超限位保持假 / Overrun stays false
    xValid := FALSE;                        // 判无效 / Invalid
    FC_DL_PreheaterStageEfficiencyCalc := FALSE;   // 返回码同步 / Return synchronised
    RETURN;                                 // 提前退出 / Early exit
END_IF

(* —— 段 3：主算式（不钳制，先出原始值供段 4 判据使用，R24） —— *)
_fDropRawK := fGasInC - fGasOutC;                                                 // 气体温降 [K]
_fApproachRawK := fGasOutC - fMatInC;                                             // 逼近温差 [K]
_fEffRawPct := _fDropRawK / _fPotentialK * DL_PCT;                                // 原始效率 [%]

(* —— 段 4：判据（取原始值；单点 BOOL 聚合避免多处赋 FALSE 覆盖） —— *)
xEffOver := (_fEffRawPct > fEffMaxPct);                                           // 超该级设计上限
xValid := (fEffMaxPct > DL_EPS)                                                   // 设计上限必须为正
          AND (fEffMaxPct <= DL_EFF_HI_PCT)                                       // 设计上限不得超过 100 %
          AND (_fEffRawPct >= DL_EFF_LO_PCT)                                      // 不低于物理域下限
          AND (_fEffRawPct <= DL_EFF_HI_PCT)                                      // 不高于物理域上限
          AND (_fDropRawK >= DL_ZERO_K)                                           // 气体必须降温（方向固定）
          AND (_fApproachRawK > DL_ZERO_K);                                       // 出口气体仍须高于进口物料

(* —— 段 5：输出单点写盘（钳制到物理域内，判定结果已在段 4 定案） —— *)
fEffPct := LIMIT(DL_EFF_LO_PCT, _fEffRawPct, DL_EFF_HI_PCT);                       // 效率钳 0..100 [%]
fGasDropK := MAX(DL_ZERO_K, _fDropRawK);                                           // 温降钳 >= 0 [K]
fApproachK := MAX(DL_ZERO_K, _fApproachRawK);                                      // 逼近温差钳 >= 0 [K]
FC_DL_PreheaterStageEfficiencyCalc := xValid;                                      // 返回码：TRUE = 计算可信

END_FUNCTION

(* ---- FC_DL_PressSectionDewaterCalc.st ---- *)
(*
  DL Factory R84 | FC_DL_PressSectionDewaterCalc
  功能：压榨部脱水，按入口干度与压榨比压、车速经验式估算出口干度与断纸风险
  开源溯源：无（clean-room 自研，依据公开工艺公式，来源=行业通用公式，许可证=MIT，借鉴点=公式结构）
  规则：R1-R16 全遵守
*)
FUNCTION FC_DL_PressSectionDewaterCalc : REAL
VAR_INPUT
    fInDryPct : REAL := 20.0; // 压榨入口干度 [%] / inlet dryness [%]
    fPressMpa : REAL := 0.8; // 压榨线比压 [MPa] / press nip line load converted to pressure [MPa]
    fSpeedMpm : REAL := 900.0; // 车速 [m/min] / machine speed [m/min]
    fGainCoefPctMpa : REAL := 8.0; // 压榨增益系数（单位比压干度提升） [%/MPa] / gain coefficient [%/MPa]
    fSpeedCoef : REAL := 0.001; // 车速衰减系数 [min/m] / speed decay coefficient [min/m]
    fDryMaxPct : REAL := 50.0; // 出口干度上限（压榨能力极限） [%] / maximum outlet dryness [%]
    fDryMinPct : REAL := 30.0; // 断纸风险干度下限 [%] / dryness floor against web breaks [%]
END_VAR
VAR_OUTPUT
    fGainPct : REAL; // 干度提升量 [%] / dryness gain [%]
    xRisk : BOOL; // 断纸风险位（出口干度低于下限） [-] / web break risk flag [-]
    xValid : BOOL; // 计算结果有效标志 [-] / calculation valid flag [-]
END_VAR
VAR
    fDen : REAL; // 车速衰减项（已加下限闸） [-] / speed decay term with a floor [-]
    fOutPct : REAL; // 出口干度中间量 [%] / outlet dryness intermediate [%]
END_VAR

// 段 1｜出口预置（R256）
FC_DL_PressSectionDewaterCalc := -1.0; // 哨兵返回 -1（无效） [-] / sentinel return -1, invalid [-]
fGainPct := 0.0; // 干度提升预置零 [%] / gain preset zero [%]
xRisk := FALSE; // 风险位预置 FALSE [-] / risk preset false [-]
xValid := FALSE; // 计算完成前不认结果 [-] / unusable before calculation [-]

// 段 2｜非有限拦截 + 域闸（R4/R20）
IF NOT (fInDryPct > -1.0E30 AND fInDryPct < 1.0E30) OR NOT (fPressMpa > -1.0E30 AND fPressMpa < 1.0E30) OR NOT (fSpeedMpm > -1.0E30 AND fSpeedMpm < 1.0E30) THEN
    RETURN; // 干度/比压/车速任一非有限即拒算 [-] / any non finite dryness, pressure or speed rejected [-]
END_IF
IF NOT (fGainCoefPctMpa > -1.0E30 AND fGainCoefPctMpa < 1.0E30) OR NOT (fSpeedCoef > -1.0E30 AND fSpeedCoef < 1.0E30) THEN
    RETURN; // 增益与衰减系数任一非有限即拒算 [-] / any non finite coefficient rejected [-]
END_IF
IF fInDryPct < 0.0 OR fInDryPct >= 100.0 OR fPressMpa < 0.0 OR fSpeedMpm < 0.0 OR fSpeedCoef < 0.0 THEN
    RETURN; // 干度开区间 + 比压与车速非负域闸 [%, MPa, m/min] / dryness open interval and non negative gate [-]
END_IF
IF fDryMaxPct < 1.0E-9 OR NOT (fDryMinPct < fDryMaxPct) THEN
    RETURN; // 干度上限正域闸 + 门限组态闸（下限须小于上限） [%] / dryness ceiling and threshold config gate [%]
END_IF

// 段 3｜经验式：增益 = k×比压 / (1 + 车速衰减项)
fDen := 1.0 + (fSpeedCoef * fSpeedMpm); // 无量纲：1 + (min/m × m/min) = - / dimensionless one plus the speed term
IF fDen < 1.0E-9 THEN
    RETURN; // 分母闸：衰减项退化 [无量纲] / denominator gate on the speed term [-]
END_IF
fGainPct := (fGainCoefPctMpa * fPressMpa) / fDen; // (%/MPa × MPa) ÷ 无量纲 = % / [%/MPa] × [MPa] / [-] = [%]
IF fGainPct < 0.0 THEN
    fGainPct := 0.0; // 负增益钳零（压榨不会使干度下降） [%] / clamp to zero, pressing never lowers dryness [%]
END_IF

// 段 4｜出口干度与上限钳位
fOutPct := fInDryPct + fGainPct; // % + % = % / [%] + [%] = [%]
IF fOutPct > fDryMaxPct THEN
    fGainPct := fDryMaxPct - fInDryPct; // 反算实际可提升量（封顶后） [%] / recompute the gain after capping [%]
    fOutPct := fDryMaxPct; // 出口干度封顶（压榨能力极限） [%] / cap the outlet dryness [%]
END_IF
IF fOutPct > 99.0 THEN
    fOutPct := 99.0; // 物理上限兜底：干度不可能达 100% [%] / physical ceiling, dryness cannot reach one hundred [%]
END_IF
IF NOT (fOutPct > -1.0E30 AND fOutPct < 1.0E30) OR NOT (fGainPct > -1.0E30 AND fGainPct < 1.0E30) THEN
    RETURN; // 结果非有限再拦一次 [-] / second finiteness gate on the results [-]
END_IF

// 段 5｜断纸风险判定：出口干度低于下限即湿部断纸风险
xRisk := fOutPct < fDryMinPct; // 直比门限，禁浮点等值 [-] / direct compare against the floor [-]
xValid := TRUE; // 链路有效 [-] / chain valid [-]
FC_DL_PressSectionDewaterCalc := fOutPct; // 返回出口干度 [%] / return the outlet dryness [%]
END_FUNCTION

(* ---- FC_DL_QuenchDelayCalc.st ---- *)
(*
  Name: FC_DL_QuenchDelayCalc
  Category: DL_Process
  Version: 1.0.0
  Round: R89 / 2026-11-25
  开源溯源：clean-room 自研（族 锻造加热退火，ST 开源生态实测 0 命中，无外部代码引入）
  功能：淬火转移延迟允许上限核算：按转移距离与速度算转移时间，估算空冷温降并判是否超允降。
  边界条件：① 四入参全部过非有限闸，任一非有限返回哨兵 -1；
            ② 转移速度为除子，按 0.05~10 m/s 域闸拦截，绝无零除；
            ③ 温降估算按空冷速率线性近似（忽略辐射非线性段），结论用于上限校核不用于工艺反算。
  量纲自证：m ÷ (m/s) = s；s × (℃/s) = ℃；与 fTempDropMaxC[℃] 同量纲比较。
*)
FUNCTION FC_DL_QuenchDelayCalc : REAL
VAR_INPUT
    fTransferDistM : REAL;      (* 转移距离（炉口至淬火槽） [m] Transfer distance [m] *)
    fTransferSpeedMps : REAL;   (* 转移机构平均速度 [m/s] Transfer speed [m/s] *)
    fTempDropMaxC : REAL;       (* 允许最大温降 [℃] Allowed maximum temperature drop [degC] *)
    fCoolRateCps : REAL;        (* 空冷速率（转移区间） [℃/s] Air cooling rate [degC/s] *)
END_VAR
VAR_OUTPUT
    fDelayS : REAL;             (* 转移时间（允许延迟上限的基准） [s] Transfer time [s] *)
    fTempDropEstC : REAL;       (* 估算温降 [℃] Estimated temperature drop [degC] *)
    xWithinLimit : BOOL;        (* 温降在允许范围内 [-] Drop within limit *)
    xValid : BOOL;              (* 计算有效性标志 [-] Calculation valid flag *)
END_VAR
VAR CONSTANT
    DL_EPS : REAL := 1.0E-9;        (* 判据容差 [-] Criterion tolerance *)
    DL_DIST_MAX : REAL := 50.0;     (* 转移距离上限 [m] Distance ceiling [m] *)
    DL_V_MIN : REAL := 0.05;        (* 转移速度下限 [m/s] Speed floor [m/s] *)
    DL_V_MAX : REAL := 10.0;        (* 转移速度上限 [m/s] Speed ceiling [m/s] *)
    DL_DROP_MIN : REAL := 5.0;      (* 允许温降下限 [℃] Drop allowance floor [degC] *)
    DL_DROP_MAX : REAL := 500.0;    (* 允许温降上限 [℃] Drop allowance ceiling [degC] *)
    DL_CR_MIN : REAL := 0.1;        (* 空冷速率下限 [℃/s] Cooling rate floor [degC/s] *)
    DL_CR_MAX : REAL := 100.0;      (* 空冷速率上限 [℃/s] Cooling rate ceiling [degC/s] *)
END_VAR
(* 出口预置：四出口统一预置（R256） *)
fDelayS := 0.0; fTempDropEstC := 0.0; xWithinLimit := FALSE; xValid := FALSE;
(* 非有限闸：NaN 自反判 + Inf 差值自减判，四入参全枚举 *)
IF (fTransferDistM <> fTransferDistM) OR ((fTransferDistM - fTransferDistM) <> 0.0)
   OR (fTransferSpeedMps <> fTransferSpeedMps) OR ((fTransferSpeedMps - fTransferSpeedMps) <> 0.0)
   OR (fTempDropMaxC <> fTempDropMaxC) OR ((fTempDropMaxC - fTempDropMaxC) <> 0.0)
   OR (fCoolRateCps <> fCoolRateCps) OR ((fCoolRateCps - fCoolRateCps) <> 0.0) THEN
    FC_DL_QuenchDelayCalc := -1.0;          (* 哨兵 -1：入参非有限 / Sentinel -1, non-finite input *)
    RETURN;
END_IF
(* 组态域闸：距离、速度为除子、允许温降、空冷速率逐项定域 *)
IF (fTransferDistM < 0.0) OR (fTransferDistM > DL_DIST_MAX)
   OR (fTransferSpeedMps < DL_V_MIN) OR (fTransferSpeedMps > DL_V_MAX)
   OR (fTempDropMaxC < DL_DROP_MIN) OR (fTempDropMaxC > DL_DROP_MAX)
   OR (fCoolRateCps < DL_CR_MIN) OR (fCoolRateCps > DL_CR_MAX) THEN
    FC_DL_QuenchDelayCalc := -1.0;          (* 哨兵 -1：组态非法 / Sentinel -1, bad configuration *)
    RETURN;
END_IF
(* 转移时间：m ÷ (m/s) = s，速度已过下限闸，绝无零除 *)
fDelayS := fTransferDistM / fTransferSpeedMps;
(* 温降估算：s × (℃/s) = ℃，线性近似（辐射非线性段由工艺余量覆盖） *)
fTempDropEstC := fDelayS * fCoolRateCps;
(* 校核：温降不超过允许值（两侧同量纲 ℃，禁浮点判等） *)
xWithinLimit := fTempDropEstC <= fTempDropMaxC;
xValid := TRUE;                             (* 链路有效 / Chain valid *)
FC_DL_QuenchDelayCalc := fDelayS;
END_FUNCTION

(* ---- FC_DL_QuenchOilTempRiseCalc.st ---- *)
(*
  Component : FC_DL_QuenchOilTempRiseCalc
  Category  : DL_Process
  Type      : FC
  Complexity: C2
  VERSION   : v1.0.0
  功能      : 淬火油槽温升与换热负荷核算：由油量/比热/工件带入热量与换热器能力算单周期温升、热平衡稳态油温与超温判定。
  开源溯源  : 道莅原创 clean-room 自研（无外部代码引用）｜License: MIT
  边界条件  : ① 油量/比热/周期时长/换热能力均须 > 1e-9，组态非法返回哨兵 -1；
              ② 稳态油温按集总热平衡估算，不含辐射与强制对流分段模型；
              ③ 超限判定用容差比较，禁浮点等值比较。
*)
FUNCTION FC_DL_QuenchOilTempRiseCalc : REAL
VAR_INPUT
    fOilMassKg  : REAL;   (* 油槽油量 [kg] Oil mass in tank *)
    fOilCpKJkgK : REAL;   (* 油比热容 [kJ/(kg·K)] Oil specific heat capacity *)
    fPartHeatKJ : REAL;   (* 单周期工件带入热量 [kJ] Heat input by parts per cycle *)
    fOilTemp0C  : REAL;   (* 初始油温 [°C] Initial oil temperature *)
    fCycleTimeS : REAL;   (* 生产周期时长 [s] Production cycle time *)
    fExchCapKWperK : REAL; (* 换热器换热能力（k·A 传导率）[kW/K] Heat exchanger conductance k*A *)
    fTempLimC   : REAL;   (* 油温允许上限 [°C] Oil temperature limit *)
END_VAR
VAR_OUTPUT
    fTempRiseK   : REAL;  (* 单周期油温升幅 [K] Temperature rise per cycle *)
    fSteadyTempC : REAL;  (* 热平衡稳态油温 [°C] Steady-state oil temperature *)
    xOverTemp    : BOOL;  (* 稳态油温超限标志 [-] Over-limit flag *)
    xValid       : BOOL;  (* 计算有效性标志 [-] Calculation valid flag *)
END_VAR
VAR CONSTANT
    DL_EPS : REAL := 1.0E-9;   (* 除零判定容差 [无量纲] Divide-by-zero tolerance *)
END_VAR
(* 出口预置：四出口统一预置，杜绝幽灵值 *)
fTempRiseK := 0.0; fSteadyTempC := 0.0; xOverTemp := FALSE; xValid := FALSE;
(* 非有限拦截：自反判 NaN，自身差值判 Inf，禁阈值近似判定 *)
IF (fOilMassKg <> fOilMassKg) OR ((fOilMassKg - fOilMassKg) <> 0.0)
   OR (fOilCpKJkgK <> fOilCpKJkgK) OR ((fOilCpKJkgK - fOilCpKJkgK) <> 0.0)
   OR (fPartHeatKJ <> fPartHeatKJ) OR ((fPartHeatKJ - fPartHeatKJ) <> 0.0)
   OR (fOilTemp0C <> fOilTemp0C) OR ((fOilTemp0C - fOilTemp0C) <> 0.0)
   OR (fCycleTimeS <> fCycleTimeS) OR ((fCycleTimeS - fCycleTimeS) <> 0.0)
   OR (fExchCapKWperK <> fExchCapKWperK) OR ((fExchCapKWperK - fExchCapKWperK) <> 0.0)
   OR (fTempLimC <> fTempLimC) OR ((fTempLimC - fTempLimC) <> 0.0) THEN
    FC_DL_QuenchOilTempRiseCalc := -1.0;   (* 哨兵 -1：输入非有限 / Sentinel -1 non-finite *)
    RETURN;
END_IF
(* 组态域闸：覆盖每一个参与判据换算的分母引脚 *)
IF (fOilMassKg <= DL_EPS) OR (fOilCpKJkgK <= DL_EPS)
   OR (fCycleTimeS <= DL_EPS) OR (fExchCapKWperK <= DL_EPS) THEN
    FC_DL_QuenchOilTempRiseCalc := -1.0;   (* 哨兵 -1：组态非法 / Sentinel -1 bad config *)
    RETURN;
END_IF
(* 单周期温升：dT = Q / (m*cp)，分母已过域闸 *)
fTempRiseK := fPartHeatKJ / (fOilMassKg * fOilCpKJkgK);
(* 热平衡稳态：热源平均功率 P = Q/t [kJ/s = kW]；稳态温升 dT = P / (k*A) [kW / (kW/K) = K]，量纲自洽 *)
fSteadyTempC := fOilTemp0C + (fPartHeatKJ / fCycleTimeS) / fExchCapKWperK;
(* 超限判定：容差比较，禁等值比较 *)
xOverTemp := fSteadyTempC > (fTempLimC + DL_EPS);
xValid := TRUE;                            (* 链路有效 / Chain valid *)
FC_DL_QuenchOilTempRiseCalc := fSteadyTempC;   (* 返回稳态油温 [°C] / Return steady temp *)
END_FUNCTION

(* ---- FC_DL_ReactorAdiabaticRise.st ---- *)
(*
  DL Factory R84 | FC_DL_ReactorAdiabaticRise
  功能：由累积投料摩尔与反应焓算绝热温升，并带投料完成度修正
  开源溯源：无（clean-room 自研，依据公开工艺公式，来源=行业通用公式，许可证=MIT，借鉴点=公式结构）
  规则：R1-R16 全遵守
*)
FUNCTION FC_DL_ReactorAdiabaticRise : REAL
VAR_INPUT
    fChargedMol : REAL := 500.0; // 已累积投料摩尔数 [mol] / charged moles so far [mol]
    fTargetMol : REAL := 800.0; // 计划满批摩尔数 [mol] / planned full batch moles [mol]
    fHrKjMol : REAL := 120.0; // 反应焓（放热取正） [kJ/mol] / heat of reaction, exotherm positive [kJ/mol]
    fMassKg : REAL := 2000.0; // 釜内物料总质量 [kg] / total batch mass [kg]
    fCpKjKgK : REAL := 3.2; // 物料比热 [kJ/(kg·K)] / batch specific heat [kJ/(kg*K)]
END_VAR
VAR_OUTPUT
    fAccumMol : REAL; // 累积投料摩尔（回显链路量） [mol] / accumulated charged moles [mol]
    fFillRatio : REAL; // 投料完成度（钳位 0~1） [-] / charge completion ratio, clamped [-]
    xValid : BOOL; // 计算结果有效标志 [-] / calculation valid flag [-]
END_VAR
VAR
    fDTadFullK : REAL; // 满批绝热温升 [K] / full batch adiabatic rise [K]
    fDTadK : REAL; // 修正后绝热温升 [K] / corrected adiabatic rise [K]
END_VAR

// 段 1｜出口预置（R256）
FC_DL_ReactorAdiabaticRise := -1.0; // 哨兵返回 -1（无效） [-] / sentinel return -1, invalid [-]
fAccumMol := 0.0; // 累积摩尔预置零 [mol] / accumulated moles preset zero [mol]
fFillRatio := 0.0; // 完成度预置零 [-] / completion preset zero [-]
xValid := FALSE; // 计算完成前不认结果 [-] / unusable before calculation [-]

// 段 2｜非有限拦截 + 域闸（R4/R20）
IF NOT (fChargedMol > -1.0E30 AND fChargedMol < 1.0E30) OR NOT (fTargetMol > -1.0E30 AND fTargetMol < 1.0E30) OR NOT (fHrKjMol > -1.0E30 AND fHrKjMol < 1.0E30) OR NOT (fMassKg > -1.0E30 AND fMassKg < 1.0E30) OR NOT (fCpKjKgK > -1.0E30 AND fCpKjKgK < 1.0E30) THEN
    RETURN; // 任一入参为 NaN/Inf 一律拒绝 [-] / any NaN or Inf input rejected [-]
END_IF
IF fTargetMol < 1.0E-9 OR fMassKg < 1.0E-9 OR fCpKjKgK < 1.0E-9 OR fChargedMol < 0.0 THEN
    RETURN; // 满批摩尔分母闸 + 质量/比热正域闸（防除零） [mol, kg] / denominator and positive domain gate [-]
END_IF

// 段 3｜满批绝热温升 ΔTad = (n·ΔHr)/(m·cp)
fDTadFullK := (fTargetMol * fHrKjMol) / (fMassKg * fCpKjKgK); // (mol × kJ/mol) ÷ (kg × kJ/(kg·K)) = K / [mol]×[kJ/mol] / ([kg]×[kJ/(kg*K)]) = [K]
IF NOT (fDTadFullK > -1.0E30 AND fDTadFullK < 1.0E30) THEN
    RETURN; // 结果非有限再拦一次 [-] / second finiteness gate [-]
END_IF

// 段 4｜投料完成度修正（钳位 0~1，超投按满批计）
fFillRatio := fChargedMol / fTargetMol; // mol ÷ mol = 无量纲 / [mol] / [mol] = [-]
IF fFillRatio > 1.0 THEN
    fFillRatio := 1.0; // 超投钳位：温升潜力按满批封顶 [-] / clamp high, potential capped at full batch [-]
END_IF
IF fFillRatio < 0.0 THEN
    fFillRatio := 0.0; // 负投料钳零 [-] / clamp low to zero [-]
END_IF
fDTadK := fDTadFullK * fFillRatio; // K × 无量纲 = K（等价于按累积摩尔计） / [K] × [-] = [K]
IF NOT (fDTadK > -1.0E30 AND fDTadK < 1.0E30) THEN
    RETURN; // 结果非有限再拦一次 [-] / second finiteness gate [-]
END_IF
fAccumMol := fChargedMol; // 回显累积投料摩尔 [mol] / echo the accumulated moles [mol]
xValid := TRUE; // 链路有效 [-] / chain valid [-]
FC_DL_ReactorAdiabaticRise := fDTadK; // 返回绝热温升 [K] / return the adiabatic rise [K]
END_FUNCTION

(* ---- FC_DL_ReactorHeatReleaseCalc.st ---- *)
(*
  DL Factory R84 | FC_DL_ReactorHeatReleaseCalc
  功能：由夹套温差流量算移热功率，叠加釜内蓄热反算放热速率与单位质量放热
  开源溯源：无（clean-room 自研，依据公开工艺公式，来源=行业通用公式，许可证=MIT，借鉴点=公式结构）
  规则：R1-R16 全遵守
*)
FUNCTION FC_DL_ReactorHeatReleaseCalc : REAL
VAR_INPUT
    fFlowKgh : REAL := 3000.0; // 夹套冷却介质流量 [kg/h] / jacket coolant flow [kg/h]
    fCpKjKgK : REAL := 4.18; // 冷却介质比热 [kJ/(kg·K)] / coolant specific heat [kJ/(kg*K)]
    fTinC : REAL := 25.0; // 夹套进口温度 [℃] / jacket inlet temperature [C]
    fToutC : REAL := 30.0; // 夹套出口温度 [℃] / jacket outlet temperature [C]
    fMassKg : REAL := 2000.0; // 釜内物料总质量 [kg] / batch mass [kg]
    fCpBatchKjKgK : REAL := 3.2; // 釜内物料比热 [kJ/(kg·K)] / batch specific heat [kJ/(kg*K)]
    fHeatRateKmin : REAL := 0.2; // 釜内温升速率 [K/min] / batch heating rate [K/min]
    fAccumKj : REAL := 1000.0; // 累计放热量 [kJ] / accumulated heat released [kJ]
END_VAR
VAR_OUTPUT
    fQremKw : REAL; // 夹套移热功率 [kW] / removed heat duty [kW]
    fQrelKjKg : REAL; // 单位质量累计放热 [kJ/kg] / specific heat released [kJ/kg]
    xValid : BOOL; // 计算结果有效标志 [-] / calculation valid flag [-]
END_VAR
VAR
    fQAccumKw : REAL; // 釜内蓄热功率 [kW] / batch accumulation duty [kW]
    fQrelKw : REAL; // 总放热速率 [kW] / total release rate [kW]
END_VAR
VAR CONSTANT
    DL_RHR_SECH : REAL := 3600.0; // 小时转秒常量 [s/h] / seconds per hour [s/h]
    DL_RHR_MIN : REAL := 60.0; // 分钟转秒常量 [s/min] / seconds per minute [s/min]
END_VAR

// 段 1｜出口预置（R256）
FC_DL_ReactorHeatReleaseCalc := -1.0; // 哨兵返回 -1（无效） [-] / sentinel return -1, invalid [-]
fQremKw := 0.0; // 移热功率预置零 [kW] / removed duty preset zero [kW]
fQrelKjKg := 0.0; // 单位放热预置零 [kJ/kg] / specific heat preset zero [kJ/kg]
xValid := FALSE; // 计算完成前不认结果 [-] / unusable before calculation [-]

// 段 2｜非有限拦截 + 域闸（R4/R20）
IF NOT (fFlowKgh > -1.0E30 AND fFlowKgh < 1.0E30) OR NOT (fCpKjKgK > -1.0E30 AND fCpKjKgK < 1.0E30) OR NOT (fTinC > -1.0E30 AND fTinC < 1.0E30) OR NOT (fToutC > -1.0E30 AND fToutC < 1.0E30) OR NOT (fMassKg > -1.0E30 AND fMassKg < 1.0E30) THEN
    RETURN; // 温度/流量/比热任一非有限即拒算 [-] / any non finite thermal input rejected [-]
END_IF
IF NOT (fCpBatchKjKgK > -1.0E30 AND fCpBatchKjKgK < 1.0E30) OR NOT (fHeatRateKmin > -1.0E30 AND fHeatRateKmin < 1.0E30) OR NOT (fAccumKj > -1.0E30 AND fAccumKj < 1.0E30) THEN
    RETURN; // 物料比热/温升速率/累积量任一非有限即拒算 [-] / any non finite batch input rejected [-]
END_IF
IF fCpKjKgK < 1.0E-9 OR fCpBatchKjKgK < 1.0E-9 OR fMassKg < 1.0E-9 OR fFlowKgh < 0.0 THEN
    RETURN; // 比热与质量正域分母闸（防除零） [kJ/(kg·K), kg] / positive cp and mass denominator gate [-]
END_IF

// 段 3｜夹套移热 Q = m·cp·ΔT（kg/s 化后即 kW）
fQremKw := (fFlowKgh / DL_RHR_SECH) * fCpKjKgK * (fToutC - fTinC); // kg/h ÷ 3600 = kg/s；kg/s × kJ/(kg·K) × K = kJ/s = kW / [kg/h] / 3600 × [kJ/(kg*K)] × [K] = [kW]
IF NOT (fQremKw > -1.0E30 AND fQremKw < 1.0E30) THEN
    RETURN; // 结果非有限再拦一次 [-] / second finiteness gate [-]
END_IF

// 段 4｜釜内蓄热功率（温升速率 K/min 化到 K/s）
fQAccumKw := (fMassKg * fCpBatchKjKgK * fHeatRateKmin) / DL_RHR_MIN; // kg × kJ/(kg·K) × K/min ÷ 60 = kJ/s = kW / [kg] × [kJ/(kg*K)] × [K/min] / 60 = [kW]

// 段 5｜总放热速率与单位质量放热
fQrelKw := fQremKw + fQAccumKw; // kW + kW = kW（放热 = 移热 + 蓄热） / [kW] + [kW] = [kW]
fQrelKjKg := fAccumKj / fMassKg; // kJ ÷ kg = kJ/kg / [kJ] / [kg] = [kJ/kg]
IF NOT (fQrelKw > -1.0E30 AND fQrelKw < 1.0E30) OR NOT (fQrelKjKg > -1.0E30 AND fQrelKjKg < 1.0E30) THEN
    RETURN; // 结果非有限再拦一次 [-] / second finiteness gate on the results [-]
END_IF
xValid := TRUE; // 链路有效 [-] / chain valid [-]
FC_DL_ReactorHeatReleaseCalc := fQrelKw; // 返回放热速率 [kW] / return the release rate [kW]
END_FUNCTION

(* ---- FC_DL_ReagentConsumeCalc.st ---- *)
(*
  道莅工业代码库 / Daoli Industrial ST Library
  组件: FC_DL_ReagentConsumeCalc
  分类: DL_Process
  开源溯源: 无（clean-room 工程公式自研；参考公开工艺计算公式，未复制任何受版权保护代码）
  许可证: 本项目自有 (MIT)
  功能: 按进出口浓度差与化学计量比折算药剂消耗速率、日耗量与药罐可用天数
*)
FUNCTION FC_DL_ReagentConsumeCalc : BOOL
VAR_INPUT
    rGasNm3h : REAL; // 标态烟气量 [Nm3/h] / flue gas flow at normal conditions
    rInMgNm3 : REAL; // 入口污染物浓度 [mg/Nm3] / inlet pollutant concentration
    rOutMgNm3 : REAL; // 出口污染物浓度 [mg/Nm3] / outlet pollutant concentration
    rStoichRatio : REAL; // 药剂与污染物的质量化学计量比 [kg/kg] / stoichiometric mass ratio
    rTankKg : REAL; // 药罐当前存量 [kg] / reagent inventory in tank
END_VAR
VAR_OUTPUT
    rKgH : REAL; // 药剂小时消耗量 [kg/h] / reagent consumption per hour
    rKgDay : REAL; // 药剂日消耗量 [kg/d] / reagent consumption per day
    rDaysLeft : REAL; // 存量可用天数 [d] / inventory remaining in days
    bValid : BOOL; // 结果有效位 [-] / result valid flag
    iErrCode : INT; // 事件码 0=正常 1=药罐存量非法 2=无脱除量无法推算天数 3=结果非有限 / event code
END_VAR
VAR CONSTANT
    rMgToKg : REAL := 1.0E-6; // 毫克转公斤系数 [kg/mg] / milligram to kilogram factor
    rHourPerDay : REAL := 24.0; // 每日小时数 [h/d] / hours per day
END_VAR
VAR
    rRemovalMgNm3 : REAL; // 净脱除浓度差 [mg/Nm3] / net removed concentration
    rKgHRaw : REAL; // 未校验小时消耗 [kg/h] / unchecked hourly consumption
END_VAR

    // —— 段 0：全路径预清 —— //
    rRemovalMgNm3 := 0.0;
    rKgHRaw := 0.0;
    rKgH := 0.0;
    rKgDay := 0.0;
    rDaysLeft := 0.0;
    bValid := FALSE;
    iErrCode := 0;
    FC_DL_ReagentConsumeCalc := FALSE;
    // —— 段 1：药罐存量域闸 —— //
    IF rTankKg <= 0.0 THEN
        iErrCode := 1; // 药罐存量非法，可用天数置零 / invalid inventory, days left zeroed
        RETURN;
    END_IF;
    // —— 段 2：量纲链 (mg/Nm3)*(Nm3/h)*(kg/mg) = kg/h；× (kg/kg) 仍为 kg/h —— //
    rRemovalMgNm3 := rInMgNm3 - rOutMgNm3; // 脱除浓度差 [mg/Nm3] / removed concentration
    IF rRemovalMgNm3 < 0.0 THEN
        rRemovalMgNm3 := 0.0; // 出口高于入口（仪表漂移）按零脱除 / outlet above inlet treated as no removal
    END_IF;
    rKgHRaw := rRemovalMgNm3 * rGasNm3h * rMgToKg * rStoichRatio; // 药剂消耗 [kg/h] / reagent consumption
    IF ABS(rKgHRaw) > 1.0E15 THEN
        iErrCode := 3; // 结果非有限，强制归零 / non-finite result, forced to zero
        RETURN;
    END_IF;
    rKgH := rKgHRaw;
    // —— 段 3：日耗量 = 小时量 × 24（量纲 kg/h × h/d = kg/d） —— //
    rKgDay := rKgH * rHourPerDay; // 日耗量 [kg/d] / daily consumption
    // —— 段 4：可用天数（分母闸：日耗必须为正） —— //
    IF rKgDay <= 1.0E-9 THEN
        iErrCode := 2; // 无脱除量，天数无法推算，置零 / no consumption, days not derivable
        bValid := TRUE;
        FC_DL_ReagentConsumeCalc := TRUE;
        RETURN;
    END_IF;
    rDaysLeft := rTankKg / rKgDay; // 可用天数 [d] / remaining days
    IF ABS(rDaysLeft) > 1.0E15 THEN
        rDaysLeft := 0.0;
        iErrCode := 3; // 结果非有限，强制归零 / non-finite result, forced to zero
        RETURN;
    END_IF;
    bValid := TRUE;
    FC_DL_ReagentConsumeCalc := TRUE;
END_FUNCTION

(* ---- FC_DL_ReceiverPressureDropCalc.st ---- *)
(*
  ============================================================
  组件名 : FC_DL_ReceiverPressureDropCalc
  分类   : DL_Process
  功能   : 储气罐压降法流量估算，由起止压力与罐容时长求标准状态流量与压降速率
  复杂度 : C1
  版本   : 1.0.0
  作者   : 道莅工业代码库工厂 / R81
  日期   : 2026-11-24
  开源溯源 : clean-room（no upstream）—— 依据公开工程公式自研，未复制任何上游实现
  红线自检 : R1 无GVL/R2 无物理地址/R3 纯IEC/R4 防除零/R5 双语注释
  接口说明 :
      标准状态流量 = (起始压力 - 终止压力) * 罐容 / 时长 * 60，单位 Nm3/min，
      该式为忽略温度补偿的工程近似，仅在罐内温度稳定且压降不超过初始压力的前提下可用。
      压降速率 = (起始压力 - 终止压力) / 时长 * 3600，单位 bar/h。
      终止压力高于起始压力表示罐在充气而非放气，本组件判为不适用并置无效。
  ============================================================
*)
FUNCTION FC_DL_ReceiverPressureDropCalc : BOOL
VAR_INPUT
    bEnable   : BOOL; // 使能：TRUE 时计算 / Enable: TRUE to compute
    bErr      : BOOL; // 外部故障：TRUE 时立即退出并置结果无效 / External fault: TRUE aborts with invalid result
    rP1_bar   : REAL; // 统计窗口起始压力 [bar] / pressure at the start of the window [bar]
    rP2_bar   : REAL; // 统计窗口终止压力 [bar] / pressure at the end of the window [bar]
    rVol_m3   : REAL; // 储气罐有效容积 [m3] / effective receiver volume [cubic metre]
    rDur_s    : REAL; // 统计窗口时长 [s] / duration of the window [second]
END_VAR
VAR_OUTPUT
    rFlow_nm3min : REAL; // 折算标准状态流量 [Nm3/min] / equivalent standard state flow [normal cubic metre per minute]
    rDropRate_barh : REAL; // 折算压降速率 [bar/h] / equivalent pressure drop rate [bar per hour]
    bValid    : BOOL; // 输出有效：TRUE 表示结果可用 / Output valid
END_VAR
VAR CONSTANT
    DL_R_MAX  : REAL := 3.0E38;  // 实数上界，用于拦截 Inf [无量纲] / real upper bound used to reject infinity [dimensionless]
    DL_EPS    : REAL := 1.0E-12; // 除零判定阈值 [无量纲] / division guard threshold [dimensionless]
    DL_S_PER_MIN : REAL := 60.0;   // 每分钟秒数 [s/min] / seconds per minute [second per minute]
    DL_S_PER_H   : REAL := 3600.0; // 每小时秒数 [s/h] / seconds per hour [second per hour]
    DL_DROP_MAX_PCT : REAL := 100.0; // 压降不得超过起始压力的百分比上限 [%] / pressure drop must not exceed this percentage of the start pressure [percent]
    DL_PCT    : REAL := 100.0;   // 百分数换算系数 [无量纲] / percentage scaling factor [dimensionless]
END_VAR
VAR
    _bFin  : BOOL := FALSE; // 输入有限性判定结果 / input finiteness verdict
    _rDrop : REAL := 0.0;   // 窗口内压降 [bar] / pressure drop inside the window [bar]
END_VAR

    // 段 1｜出口预置
    rFlow_nm3min := 0.0;
    rDropRate_barh := 0.0;
    bValid := FALSE;
    // 段 2｜使能闸与外部故障闸
    IF NOT bEnable THEN
        RETURN;
    END_IF;
    IF bErr THEN
        RETURN;
    END_IF;
    // 段 3｜非有限闸
    _bFin := (rP1_bar = rP1_bar) AND (ABS(rP1_bar) <= DL_R_MAX) AND (rP2_bar = rP2_bar) AND (ABS(rP2_bar) <= DL_R_MAX) AND (rVol_m3 = rVol_m3) AND (ABS(rVol_m3) <= DL_R_MAX) AND (rDur_s = rDur_s) AND (ABS(rDur_s) <= DL_R_MAX);
    IF NOT _bFin THEN
        RETURN;
    END_IF;
    // 段 4｜域闸：罐容与时长必须严格为正，压力不得为负
    IF (ABS(rVol_m3) <= DL_EPS) OR (ABS(rDur_s) <= DL_EPS) THEN
        RETURN;
    END_IF;
    IF (rVol_m3 < 0.0) OR (rDur_s < 0.0) OR (rP1_bar < 0.0) OR (rP2_bar < 0.0) THEN
        RETURN;
    END_IF;
    // 段 5｜压降必须为正，否则属充气工况，压降法不适用
    _rDrop := rP1_bar - rP2_bar;
    IF _rDrop <= DL_EPS THEN
        RETURN;
    END_IF;
    // 段 6｜压降相对起始压力不得越界，否则近似式失真
    IF rP1_bar > DL_EPS THEN
        IF _rDrop > rP1_bar * DL_DROP_MAX_PCT / DL_PCT THEN
            RETURN;
        END_IF;
    END_IF;
    // 段 7｜流量与压降速率
    rFlow_nm3min := _rDrop * rVol_m3 / rDur_s * DL_S_PER_MIN;
    rDropRate_barh := _rDrop / rDur_s * DL_S_PER_H;
    bValid := TRUE;
    FC_DL_ReceiverPressureDropCalc := bValid;
END_FUNCTION

(* ---- FC_DL_ReExtractionFactorCalc.st ---- *)
(*
  Component : FC_DL_ReExtractionFactorCalc
  Category  : DL_Process
  Function  : 稀土溶剂萃取分配比 D 与单级萃取率 E 换算，E = D / (D + O/A)
  Complexity: C2
  开源溯源 : DLF 内部原创（R94 族模板派生）；参考语义来源见 SOURCE_HUNTING_MATRIX.md
  规则遵从 : R1-R16
  契约     : 输入 rDistCoefD 分配比 [-]，rRatioOA 相比 O/A [-]；输出 rExtractFrac 萃取率 [0~1]、
             rExtractPct 萃取率 [%]、xValid 有效标志、nFaultCode 故障码；返回 TRUE 表示两输出可信。
  边界     : 分配比须 ≥0、相比须 >0；分母 D+O/A 绝对值 <1.0E-9 判 9802；任一浮点输入非有限判 9801；
             无除法以外的失效面，零全局、零物理地址、零库件依赖。
  码位     : 9801 输入非法（故障级）；9802 分母过小（故障级）。二者不并存，9801 先判。
*)
FUNCTION FC_DL_ReExtractionFactorCalc : BOOL
VAR_INPUT
    rDistCoefD : LREAL := 1.0;        // 分配比 D，有机相稀土浓度与水相稀土浓度之比 [-] EN: distribution ratio D of organic to aqueous rare earth concentration
    rRatioOA   : LREAL := 1.0;        // 相比 O/A，有机相体积流量与水相体积流量之比 [-] EN: organic to aqueous volumetric phase ratio O over A
END_VAR
VAR_OUTPUT
    rExtractFrac : LREAL;             // 单级萃取率 E 的无量纲值，域 0~1 [-] EN: single stage extraction fraction within the range zero to one
    rExtractPct  : LREAL;             // 单级萃取率 E 的百分数 [%] EN: single stage extraction efficiency expressed in percent
    xValid       : BOOL;              // 两输出可信标志 EN: both outputs are valid
    nFaultCode   : INT;               // 0=无故障 9801=分配比或相比非法 9802=分母过小 EN: zero none, 9801 illegal input, 9802 denominator too small
END_VAR
VAR
    xFinD  : BOOL;                    // 分配比有限性 EN: the distribution ratio is finite
    xFinOA : BOOL;                    // 相比有限性 EN: the phase ratio is finite
    xFinAll: BOOL;                    // 两输入同时有限 EN: both inputs are finite at the same time
    rDen   : LREAL;                   // 萃取率分母 D + O/A [-1] EN: the denominator of the extraction rate
    rFrac  : LREAL;                   // 萃取率中间值，钳位后写入出口 [-] EN: the interim extraction fraction before clamping
END_VAR
VAR CONSTANT
    DL_REF_Z       : LREAL := 0.0;    // 浮点零常量 EN: the floating point zero constant
    DL_REF_ONE     : LREAL := 1.0;    // 浮点壹常量 EN: the floating point one constant
    DL_REF_HUNDRED : LREAL := 100.0;  // 百分数换算系数 EN: the percent conversion factor
    DL_REF_DEN_MIN : LREAL := 1.0E-9; // 分母绝对值下限 EN: the lower bound of the denominator magnitude
    DL_REF_C_BAD   : INT := 9801;     // 分配比或相比非法 EN: illegal distribution ratio or phase ratio
    DL_REF_C_DEN   : INT := 9802;     // 分母过小不可除 EN: the denominator is too small to divide
END_VAR

// 段1｜出口预置：函数名即返回值，先置假与哨兵零，任何早退分支都停在此状态
FC_DL_ReExtractionFactorCalc := FALSE;   // 返回值预置假 EN: preset the return value to false
rExtractFrac := DL_REF_Z;                // 萃取率预置零 [0~1] EN: preset the extraction fraction to zero
rExtractPct := DL_REF_Z;                 // 萃取率百分数预置零 [%] EN: preset the extraction percent to zero
xValid := FALSE;                         // 有效标志预置假 EN: preset the validity flag to false
nFaultCode := 0;                         // 故障码预置零 EN: preset the fault code to zero

// 段2｜非有限闸：NaN 用自反判、Inf 用差值自减判，两输入全部列入闸内
xFinD := (rDistCoefD = rDistCoefD) AND ((rDistCoefD - rDistCoefD) = DL_REF_Z);   // 分配比有限性 EN: the distribution ratio is finite
xFinOA := (rRatioOA = rRatioOA) AND ((rRatioOA - rRatioOA) = DL_REF_Z);           // 相比有限性 EN: the phase ratio is finite
xFinAll := xFinD AND xFinOA;                                                     // 合并有限性 EN: the combined finiteness
IF NOT xFinAll THEN                                                              // 非有限直接出口 EN: leave early on a non finite input
    nFaultCode := DL_REF_C_BAD;                                                  // 输入非法码 EN: the illegal input code
    RETURN;                                                                      // 早退：出口保持预置值 EN: return early, the outputs keep the preset values
END_IF

// 段3｜域闸：分配比非负、相比为正，否则物理上无意义
IF (rDistCoefD < DL_REF_Z) OR (rRatioOA <= DL_REF_Z) THEN                        // 域闸：负分配比或非正相比 EN: a negative distribution ratio or a non positive phase ratio
    nFaultCode := DL_REF_C_BAD;                                                  // 输入非法码 EN: the illegal input code
    RETURN;                                                                      // 早退 EN: return early
END_IF

// 段4｜分母下限保护：分母由两项正量相加，仍按绝对值下限硬校验防浮点下溢
rDen := rDistCoefD + rRatioOA;                                                   // 组成萃取率分母 [-] EN: build the denominator of the extraction rate
IF ABS(rDen) < DL_REF_DEN_MIN THEN                                               // 分母下限判据 EN: the denominator magnitude gate
    nFaultCode := DL_REF_C_DEN;                                                  // 分母过小码 EN: the denominator too small code
    RETURN;                                                                      // 早退 EN: return early
END_IF

// 段5｜主体换算：E = D / (D + O/A)，两输出同一来源，避免名实不一致
rFrac := rDistCoefD / rDen;                                                      // 计算萃取率 [-] EN: compute the extraction fraction
IF rFrac < DL_REF_Z THEN                                                         // 钳位下界（仅防御浮点残差） EN: clamp the lower bound against a residual sign error
    rFrac := DL_REF_Z;                                                           // 钳到零 EN: clamp to zero
END_IF
IF rFrac > DL_REF_ONE THEN                                                       // 钳位上界 EN: clamp the upper bound
    rFrac := DL_REF_ONE;                                                         // 钳到壹 EN: clamp to one
END_IF
rExtractFrac := rFrac;                                                           // 无量纲出口 [-] EN: the dimensionless output
rExtractPct := rFrac * DL_REF_HUNDRED;                                           // 百分数出口 [%] EN: the percent output
xValid := TRUE;                                                                  // 结果可信 EN: the results are valid
nFaultCode := 0;                                                                 // 无故障 EN: no fault
FC_DL_ReExtractionFactorCalc := TRUE;                                            // 返回真 EN: return true
END_FUNCTION

(* ---- FC_DL_RefinerFreenessCalc.st ---- *)
(*
  DL Factory R84 | FC_DL_RefinerFreenessCalc
  功能：由比边缘负荷与比能耗线性估算打浆度 CSF 并给目标偏差
  开源溯源：无（clean-room 自研，依据公开工艺公式，来源=行业通用公式，许可证=MIT，借鉴点=公式结构）
  规则：R1-R16 全遵守
*)
FUNCTION FC_DL_RefinerFreenessCalc : REAL
VAR_INPUT
    fEdgeLoadJm : REAL := 1.2; // 比边缘负荷实测值 [J/m] / measured specific edge load [J/m]
    fSecKwhT : REAL := 120.0; // 比能耗 [kWh/t] / specific energy consumption [kWh/t]
    fCsfBaseMl : REAL := 650.0; // 基准打浆度（未打浆） [mL] / base freeness [mL]
    fKEffJm : REAL := 30.0; // 比边缘负荷影响系数 [mL·m/J] / edge load sensitivity [mL*m/J]
    fKEffKwhT : REAL := 0.6; // 比能耗影响系数 [mL/(kWh/t)] / energy sensitivity [mL/(kWh/t)]
    fCsfMinMl : REAL := 100.0; // 打浆度下限（钳位） [mL] / lower clamp [mL]
    fCsfMaxMl : REAL := 750.0; // 打浆度上限（钳位） [mL] / upper clamp [mL]
    fCsfTargetMl : REAL := 350.0; // 目标打浆度 [mL] / target freeness [mL]
END_VAR
VAR_OUTPUT
    fSelJm : REAL; // 比边缘负荷回显（链路校验） [J/m] / specific edge load echo [J/m]
    fDevMl : REAL; // 与目标打浆度偏差 [mL] / deviation from the target [mL]
    xValid : BOOL; // 计算结果有效标志 [-] / calculation valid flag [-]
END_VAR
VAR
    fCsfRawMl : REAL; // 未钳位估算打浆度 [mL] / unclamped freeness estimate [mL]
    fCsfMl : REAL; // 钳位后打浆度 [mL] / clamped freeness [mL]
END_VAR

// 段 1｜出口预置（R256）
FC_DL_RefinerFreenessCalc := -1.0; // 哨兵返回 -1（无效） [-] / sentinel return -1, invalid [-]
fSelJm := 0.0; // 负荷回显预置零 [J/m] / load echo preset zero [J/m]
fDevMl := 0.0; // 偏差预置零 [mL] / deviation preset zero [mL]
xValid := FALSE; // 计算完成前不认结果 [-] / unusable before calculation [-]

// 段 2｜非有限拦截 + 域闸（R4/R20）
IF NOT (fEdgeLoadJm > -1.0E30 AND fEdgeLoadJm < 1.0E30) OR NOT (fSecKwhT > -1.0E30 AND fSecKwhT < 1.0E30) OR NOT (fCsfBaseMl > -1.0E30 AND fCsfBaseMl < 1.0E30) THEN
    RETURN; // 负荷/能耗/基准值任一非有限即拒算 [-] / any non finite load, energy or base rejected [-]
END_IF
IF NOT (fKEffJm > -1.0E30 AND fKEffJm < 1.0E30) OR NOT (fKEffKwhT > -1.0E30 AND fKEffKwhT < 1.0E30) OR NOT (fCsfTargetMl > -1.0E30 AND fCsfTargetMl < 1.0E30) THEN
    RETURN; // 系数与目标值任一非有限即拒算 [-] / any non finite coefficient or target rejected [-]
END_IF
IF fEdgeLoadJm < 0.0 OR fSecKwhT < 0.0 OR fCsfBaseMl <= 0.0 OR fCsfTargetMl < 0.0 THEN
    RETURN; // 负荷/能耗非负 + 基准与目标正域闸 [J/m, kWh/t, mL] / non negative load and positive base gate [-]
END_IF
IF NOT (fCsfMinMl < fCsfMaxMl) THEN
    RETURN; // 钳位区间组态闸：下限必须严格小于上限 [mL] / clamp band config gate [mL]
END_IF

// 段 3｜线性估算：CSF = 基准 − k1×SEL − k2×SEC
fCsfRawMl := (fCsfBaseMl - (fKEffJm * fEdgeLoadJm)) - (fKEffKwhT * fSecKwhT); // mL − (mL·m/J × J/m) − (mL/(kWh/t) × kWh/t) = mL / [mL] terms subtracted, result in [mL]
IF NOT (fCsfRawMl > -1.0E30 AND fCsfRawMl < 1.0E30) THEN
    RETURN; // 结果非有限再拦一次 [-] / second finiteness gate [-]
END_IF

// 段 4｜上下限钳位（线性近似仅在工艺区间内可信）
fCsfMl := fCsfRawMl; // 先接未钳位值 [mL] / take the raw estimate [mL]
IF fCsfMl > fCsfMaxMl THEN
    fCsfMl := fCsfMaxMl; // 上限钳位：过度打浆不成立 [mL] / clamp high, over refining is not physical [mL]
END_IF
IF fCsfMl < fCsfMinMl THEN
    fCsfMl := fCsfMinMl; // 下限钳位：湿重打浆极限 [mL] / clamp low, wet freeness floor [mL]
END_IF

// 段 5｜偏差与出口
fDevMl := fCsfMl - fCsfTargetMl; // mL − mL = mL / [mL] minus [mL] = [mL]
IF NOT (fDevMl > -1.0E30 AND fDevMl < 1.0E30) THEN
    RETURN; // 结果非有限再拦一次 [-] / second finiteness gate [-]
END_IF
fSelJm := fEdgeLoadJm; // 回显实测比边缘负荷 [J/m] / echo the measured edge load [J/m]
xValid := TRUE; // 链路有效 [-] / chain valid [-]
FC_DL_RefinerFreenessCalc := fCsfMl; // 返回打浆度 [mL] / return the freeness [mL]
END_FUNCTION
